          // fill telegramm header - just for later debugging ( the header is part of the command payload itselfy ) {{{
          Telegram.PlcToRob.Sequence[_seqIdx].Fragment[_fragIdx].Command.Header.CmdType       := CombineBytesToUint ( AxesGroup.Acyclic.ActiveCommandRegister.Register[_regIdx].Command[ACTIVE_CMD].Payload[0],
                                                                                                                      AxesGroup.Acyclic.ActiveCommandRegister.Register[_regIdx].Command[ACTIVE_CMD].Payload[1]);
          Telegram.PlcToRob.Sequence[_seqIdx].Fragment[_fragIdx].Command.Header.ExecMode.0    :=                      AxesGroup.Acyclic.ActiveCommandRegister.Register[_regIdx].Command[ACTIVE_CMD].Payload[2].0;
          Telegram.PlcToRob.Sequence[_seqIdx].Fragment[_fragIdx].Command.Header.ExecMode.1    :=                      AxesGroup.Acyclic.ActiveCommandRegister.Register[_regIdx].Command[ACTIVE_CMD].Payload[2].1;
          Telegram.PlcToRob.Sequence[_seqIdx].Fragment[_fragIdx].Command.Header.ExecMode.2    :=                      AxesGroup.Acyclic.ActiveCommandRegister.Register[_regIdx].Command[ACTIVE_CMD].Payload[2].2;
          Telegram.PlcToRob.Sequence[_seqIdx].Fragment[_fragIdx].Command.Header.ExecMode.3    :=                      AxesGroup.Acyclic.ActiveCommandRegister.Register[_regIdx].Command[ACTIVE_CMD].Payload[2].3;
          Telegram.PlcToRob.Sequence[_seqIdx].Fragment[_fragIdx].Command.Header.Prio.0        :=                      AxesGroup.Acyclic.ActiveCommandRegister.Register[_regIdx].Command[ACTIVE_CMD].Payload[3].0;
          Telegram.PlcToRob.Sequence[_seqIdx].Fragment[_fragIdx].Command.Header.Prio.1        :=                      AxesGroup.Acyclic.ActiveCommandRegister.Register[_regIdx].Command[ACTIVE_CMD].Payload[3].1;
          Telegram.PlcToRob.Sequence[_seqIdx].Fragment[_fragIdx].Command.Header.Prio.2        :=                      AxesGroup.Acyclic.ActiveCommandRegister.Register[_regIdx].Command[ACTIVE_CMD].Payload[3].2;
          Telegram.PlcToRob.Sequence[_seqIdx].Fragment[_fragIdx].Command.Header.Prio.3        :=                      AxesGroup.Acyclic.ActiveCommandRegister.Register[_regIdx].Command[ACTIVE_CMD].Payload[3].3;
          Telegram.PlcToRob.Sequence[_seqIdx].Fragment[_fragIdx].Command.Header.ParSequence.0 :=                      AxesGroup.Acyclic.ActiveCommandRegister.Register[_regIdx].Command[ACTIVE_CMD].Payload[3].4;
          Telegram.PlcToRob.Sequence[_seqIdx].Fragment[_fragIdx].Command.Header.ParSequence.1 :=                      AxesGroup.Acyclic.ActiveCommandRegister.Register[_regIdx].Command[ACTIVE_CMD].Payload[3].5;
          Telegram.PlcToRob.Sequence[_seqIdx].Fragment[_fragIdx].Command.Header.ParSequence.2 :=                      AxesGroup.Acyclic.ActiveCommandRegister.Register[_regIdx].Command[ACTIVE_CMD].Payload[3].6;
          Telegram.PlcToRob.Sequence[_seqIdx].Fragment[_fragIdx].Command.Header.ParSequence.3 :=                      AxesGroup.Acyclic.ActiveCommandRegister.Register[_regIdx].Command[ACTIVE_CMD].Payload[3].7;
          // }}}
          // loop through the payload
          FOR _payLoadPtr := AxesGroup.Acyclic.ActiveCommandRegister.Register[_regIdx].Command[ACTIVE_CMD].PayLoadPtr TO AxesGroup.Acyclic.ActiveCommandRegister.Register[_regIdx].Command[ACTIVE_CMD].PayloadLen -1  
          DO
            // copy payload
            Telegram.PlcToRob.Sequence[_seqIdx].Fragment[_fragIdx].Command.Payload[_payLoadPtr] 
              := AxesGroup.Acyclic.ActiveCommandRegister.Register[_regIdx].Command[ACTIVE_CMD].Payload[_payLoadPtr];
        
            // inc current sequence payload length
            Telegram.PlcToRob.Sequence[_seqIdx].Header.PayloadLength
              := Telegram.PlcToRob.Sequence[_seqIdx].Header.PayloadLength + 1;  
        
            // inc current fragment payload length
            Telegram.PlcToRob.Sequence[_seqIdx].Fragment[_fragIdx].Header.PayloadLength 
              := Telegram.PlcToRob.Sequence[_seqIdx].Fragment[_fragIdx].Header.PayloadLength + 1;
        
            // inc payload pointer in active command register
            AxesGroup.Acyclic.ActiveCommandRegister.Register[_regIdx].Command[ACTIVE_CMD].PayLoadPtr 
              := AxesGroup.Acyclic.ActiveCommandRegister.Register[_regIdx].Command[ACTIVE_CMD].PayLoadPtr + 1;
          
            // set command state
            IF ( AxesGroup.Acyclic.ActiveCommandRegister.Register[_regIdx].Command[ACTIVE_CMD].PayLoadPtr >= AxesGroup.Acyclic.ActiveCommandRegister.Register[_regIdx].Command[ACTIVE_CMD].PayLoadLen) 
            THEN
              AxesGroup.Acyclic.ActiveCommandRegister.Register[_regIdx].Command[ACTIVE_CMD].State := BufferStateCmd.PROCESSED;
            ELSE
              AxesGroup.Acyclic.ActiveCommandRegister.Register[_regIdx].Command[ACTIVE_CMD].State := BufferStateCmd.SENDING;  
            END_IF 
    
            // calc current telegram payload length
           _telegramLengthCurrent := 4 + Telegram.PlcToRob.Sequence[_seqIdx].Header.PayloadLength; // ST-FIX F63: sequence header + payload
      
            // check limit reached ?
            IF ( _telegramLengthCurrent >= SEQUENCE_MAX_PAYLOAD_SIZE (* ST-FIX F63 *)) 
            THEN  
              EXIT; // -> abort for loop 
            END_IF  
          END_FOR
    
          // check payload complete ?
         _fragmentAction.Complete := AxesGroup.Acyclic.ActiveCommandRegister.Register[_regIdx].Command[ACTIVE_CMD].PayLoadPtr 
                                  >= AxesGroup.Acyclic.ActiveCommandRegister.Register[_regIdx].Command[ACTIVE_CMD].PayloadLen;
    
          // just for brakepoint
          IF (_fragmentAction.Complete)
          THEN
           _fragmentAction.Complete := _fragmentAction.Complete; 
          END_IF
    
          // set fragment action
          Telegram.PlcToRob.Sequence[_seqIdx].Fragment[_fragIdx].Header.FragmentAction := FragmentActionToByte(_fragmentAction);
        END_IF
      END_IF
      
      // inc execution order list index 
     _listIdx := _listIdx + 1;
      // inc fragment index 
     _fragIdx := _fragIdx + 1;
  
      // check abort conditions
      IF (( _telegramLengthCurrent                                                >= SEQUENCE_MAX_PAYLOAD_SIZE (* ST-FIX F63 *)  ) OR  // Payload limit reached 
          ( _fragIdx                                                              >=  RobotLibraryParameter.FRAGMENT_MAX ) OR  // Max fragment limit reached
          (  AxesGroup.Acyclic.ActiveCommandRegister.ExecutionOrderList[_listIdx]  =  EMPTY_EOL_ENTRY                    ))    // No entry in ExecutionOrderList left
      THEN
        EXIT;// -> Abort while loop
      END_IF         
    END_WHILE  
    
    AxesGroup.State.SequenceCountSend          := _seqCount; // ST-FIX F63
    AxesGroup.State.FragmentCountSend[_seqIdx] := _fragIdx;
    
  END_IF  
END_FOR
                
                
END_METHOD

METHOD CalculateCyclicDataLength : UINT
VAR_IN_OUT
  /// Robot assignment of function
  AxesGroup : AxesGroup;
END_VAR
VAR_INPUT
  /// Communication direction
  Direction : ComDirection;
END_VAR

VAR CONSTANT
  /// Size of the header
  ROB_TO_PLC_HEADER_SIZE : UINT := 10;
END_VAR
                  // ------------------------------------
// PLC -> ROB
// ------------------------------------
IF (Direction = ComDirection.PLC_TO_ROB)
THEN  
  // Add Header size 
  CalculateCyclicDataLength := CalculateCyclicDataLength + SIZEOF(Telegram.PlcToRob.Header);  
  // Add Cyclic size (ST-FIX F2: only with Cartesian Position RC -> PLC)
  IF ( AxesGroup.CyclicOptional.RobToPlc.CartesianPosition.Active )
  THEN
    CalculateCyclicDataLength := CalculateCyclicDataLength + SIZEOF(Telegram.PlcToRob.Cyclic);
  END_IF
  
  // Check SubProgramData active ? 
  IF ( AxesGroup.CyclicOptional.PlcToRob.SubProgramData.Active )
  THEN
    // Add SubProgramData size 
    CalculateCyclicDataLength := CalculateCyclicDataLength + SIZEOF(Telegram.PlcToRob.CyclicOptional.SubProgramData);
  END_IF
    
  // Check CartesianPosition active ? 
  IF ( AxesGroup.CyclicOptional.PlcToRob.CartesianPosition.Active )
  THEN
    // Add CartesianPosition size 
    CalculateCyclicDataLength := CalculateCyclicDataLength + SIZEOF(Telegram.PlcToRob.CyclicOptional.CartesianPosition);
  END_IF
  
  // Check JointPosition active ? 
  IF ( AxesGroup.CyclicOptional.PlcToRob.JointPosition.Active )
  THEN
    // Add JointPosition size 
    CalculateCyclicDataLength := CalculateCyclicDataLength + SIZEOF(Telegram.PlcToRob.CyclicOptional.JointPosition);
  END_IF  
  
  // Check Force active ? 
  IF ( AxesGroup.CyclicOptional.PlcToRob.Force.Active )
  THEN
    // Add Force size 
    CalculateCyclicDataLength := CalculateCyclicDataLength + SIZEOF(Telegram.PlcToRob.CyclicOptional.Force);
  END_IF  
    
  // Check CartesianPositionExt acive ? 
  IF ( AxesGroup.CyclicOptional.PlcToRob.CartesianPositionExt.Active )
  THEN
    // Add CartesianPositionExt size 
    CalculateCyclicDataLength := CalculateCyclicDataLength + SIZEOF(Telegram.PlcToRob.CyclicOptional.CartesianPositionExt);
  END_IF   
    
  // Check JointPositionExt active ?
  IF ( AxesGroup.CyclicOptional.PlcToRob.JointPositionExt.Active )
  THEN
    // Add JointPositionExt size 
    CalculateCyclicDataLength := CalculateCyclicDataLength + SIZEOF(Telegram.PlcToRob.CyclicOptional.JointPositionExt);
  END_IF  
        
  // Check ForceExt active ?
  IF ( AxesGroup.CyclicOptional.PlcToRob.ForceExt.Active )
  THEN
    // Add ForceExt size 
    CalculateCyclicDataLength := CalculateCyclicDataLength + SIZEOF(Telegram.PlcToRob.CyclicOptional.ForceExt);
  END_IF
END_IF

// ------------------------------------
// ROB -> PLC
// ------------------------------------
IF (Direction = ComDirection.ROB_TO_PLC)
THEN
  // Add Header size 
  CalculateCyclicDataLength := CalculateCyclicDataLength + ROB_TO_PLC_HEADER_SIZE; 
  // a constant, because SIZEOF(Telegram.RobToPlc.Header) counts the VersionStruct instead of one byte
  
  // Check SubProgramData active ? 
  IF ( AxesGroup.CyclicOptional.RobToPlc.SubProgramData.Active )
  THEN
    // Add SubProgramData size 
    CalculateCyclicDataLength := CalculateCyclicDataLength + SIZEOF(Telegram.RobToPlc.CyclicOptional.SubProgramData);
  END_IF
    
  // Check CartesianPosition active ? 
  IF ( AxesGroup.CyclicOptional.RobToPlc.CartesianPosition.Active )
  THEN
    // Add CartesianPosition size 
    CalculateCyclicDataLength := CalculateCyclicDataLength + SIZEOF(Telegram.RobToPlc.CyclicOptional.CartesianPosition);
  END_IF
  
  // Check JointPosition active ? 
  IF ( AxesGroup.CyclicOptional.RobToPlc.JointPosition.Active )
  THEN
    // Add JointPosition size 
    CalculateCyclicDataLength := CalculateCyclicDataLength + SIZEOF(Telegram.RobToPlc.CyclicOptional.JointPosition);
  END_IF  
  
  // Check Force active ? 
  IF ( AxesGroup.CyclicOptional.RobToPlc.Force.Active )
  THEN
    // Add Force size 
    CalculateCyclicDataLength := CalculateCyclicDataLength + SIZEOF(Telegram.RobToPlc.CyclicOptional.Force);
  END_IF  
    
  // Check Current acive ? 
  IF ( AxesGroup.CyclicOptional.RobToPlc.Current.Active )
  THEN
    // Add Current size 
    CalculateCyclicDataLength := CalculateCyclicDataLength + SIZEOF(Telegram.RobToPlc.CyclicOptional.Current);
  END_IF    
    
  // Check CartesianPositionExt acive ? 
  IF ( AxesGroup.CyclicOptional.RobToPlc.CartesianPositionExt.Active )
  THEN
    // Add CartesianPositionExt size 
    CalculateCyclicDataLength := CalculateCyclicDataLength + SIZEOF(Telegram.RobToPlc.CyclicOptional.CartesianPositionExt);
  END_IF  
    
  // Check JointPositionExt active ?
  IF ( AxesGroup.CyclicOptional.RobToPlc.JointPositionExt.Active )
  THEN
    // Add JointPositionExt size 
    CalculateCyclicDataLength := CalculateCyclicDataLength + SIZEOF(Telegram.RobToPlc.CyclicOptional.JointPositionExt);
  END_IF  
        
  // Check ForceExt active ?
  IF ( AxesGroup.CyclicOptional.RobToPlc.ForceExt.Active )
  THEN
    // Add ForceExt size 
    CalculateCyclicDataLength := CalculateCyclicDataLength + SIZEOF(Telegram.RobToPlc.CyclicOptional.ForceExt);
  END_IF
    
  // Check CurrentExt active ? 
  IF ( AxesGroup.CyclicOptional.RobToPlc.CurrentExt.Active )
  THEN
    // Add CurrentExt size 
    CalculateCyclicDataLength := CalculateCyclicDataLength + SIZEOF(Telegram.RobToPlc.CyclicOptional.CurrentExt);
  END_IF
END_IF
                
END_METHOD

METHOD CalculateSequencePayloadMax : UINT
VAR_IN_OUT
  /// Robot assignment of function
  AxesGroup : AxesGroup;
END_VAR
VAR_INPUT
  /// Communication direction
  Direction : ComDirection;
  /// Sequeunce
  Sequence : SequenceFlag;  
END_VAR

VAR
  /// Length of the cyclic header
 _cyclicDataLength      : UINT;
  /// Acyclic area (ST-FIX F63)
 _area                  : UDINT;
END_VAR
                  // calculate cyclic header length
_cyclicDataLength := CalculateCyclicDataLength(AxesGroup := AxesGroup, Direction := Direction);


// ST-FIX F63: acyclic area without the footer, halved for two sequences (spec Fig. 5-205)
IF ( Direction = ComDirection.PLC_TO_ROB )
THEN
  _area := UINT_TO_UDINT(_parCfg.Com.TelegramLengthPlcToRob) - UINT_TO_UDINT(_cyclicDataLength) - FOOTER_SIZE;
ELSE
  _area := UINT_TO_UDINT(_parCfg.Com.TelegramLengthRobToPlc) - UINT_TO_UDINT(_cyclicDataLength) - FOOTER_SIZE;
END_IF

IF ( NOT _parCfg.Com.TwoSequences )
THEN
  IF ( Sequence = SequenceFlag.PRIMARY_SEQUENCE )
  THEN
    CalculateSequencePayloadMax := UDINT_TO_UINT(_area);
  ELSE
    CalculateSequencePayloadMax := 0;
  END_IF
ELSIF ( Sequence = SequenceFlag.PRIMARY_SEQUENCE )
THEN
  CalculateSequencePayloadMax := UDINT_TO_UINT(_area / 2);
ELSE
  CalculateSequencePayloadMax := UDINT_TO_UINT(_area - _area / 2);
END_IF
                
END_METHOD

METHOD CalculateSequencePayloadStartAdr : UINT
VAR_IN_OUT
  /// Robot assignment of function
  AxesGroup : AxesGroup;
END_VAR
VAR_INPUT
  /// Communication direction
  Direction : ComDirection;
  /// Sequeunce
  Sequence : SequenceFlag;  
END_VAR

VAR
  /// Length of the cyclic header
 _cyclicDataLength      : UINT;
  /// Length of the sequnce payload
 _sequencePayloadLength : UINT;
END_VAR
                  // calculate cyclic header length
_cyclicDataLength := CalculateCyclicDataLength(AxesGroup := AxesGroup, Direction := Direction);

CASE (Sequence) 
OF

  SequenceFlag.PRIMARY_SEQUENCE   : 
  
    // return start address
    CalculateSequencePayloadStartAdr := _cyclicDataLength;

  SequenceFlag.SECONDARY_SEQUENCE :
  
    // calculate sequence payload max
   _sequencePayloadLength 
     := CalculateSequencePayloadMax( AxesGroup := AxesGroup, 
                                     Direction := Direction, 
                                     Sequence  := SequenceFlag.PRIMARY_SEQUENCE ); // ST-FIX F63: behind the area of the 1st sequence
                                     
    // return start address
    CalculateSequencePayloadStartAdr := _cyclicDataLength + _sequencePayloadLength;
    
END_CASE
                
END_METHOD

METHOD PROTECTED CalculateTelegramLengthPlcToRob : UINT
VAR_IN_OUT
  /// Robot assignment of function
  AxesGroup : AxesGroup;
END_VAR
VAR
  /// length of the cyclic data block
 _cyclicDataLength : UINT;
END_VAR
                  _cyclicDataLength := CalculateCyclicDataLength(AxesGroup := AxesGroup, Direction := ComDirection.PLC_TO_ROB); 


IF ( _parCfg.Com.TwoSequences )
THEN
  CalculateTelegramLengthPlcToRob := _cyclicDataLength
                                    + SIZEOF(Telegram.PlcToRob.Sequence[  PRIMARY_SEQUENCE].Header)
                                    +       (Telegram.PlcToRob.Sequence[  PRIMARY_SEQUENCE].Header.PayloadLength)
                                    + SIZEOF(Telegram.PlcToRob.Sequence[SECONDARY_SEQUENCE].Header)
                                    +       (Telegram.PlcToRob.Sequence[SECONDARY_SEQUENCE].Header.PayloadLength)
                                    + SIZEOF(Telegram.PlcToRob.Footer);  
ELSE
  CalculateTelegramLengthPlcToRob := _cyclicDataLength
                                    + SIZEOF(Telegram.PlcToRob.Sequence[PRIMARY_SEQUENCE].Header)
                                    +       (Telegram.PlcToRob.Sequence[PRIMARY_SEQUENCE].Header.PayloadLength)
                                    + SIZEOF(Telegram.PlcToRob.Footer);
END_IF
                
END_METHOD

/// ST-FIX F132: checks that the AxesGroup and the telegram buffers are not used by another RobotTask
/// (table 7-1: 16#8007 ERR_AXESGROUP_INVALID, 16#8008 ERR_PERIPHERY_INVALID) and registers them
METHOD PRIVATE CheckAssignmentValid : BOOL
VAR_IN_OUT
  /// Robot assignment of function
  AxesGroup    : AxesGroup;
  /// Inputs of PLC for communication from RC
  RobotInData  : ARRAY[*] OF BYTE;
  /// Outputs of PLC for communication to RC
  RobotOutData : ARRAY[*] OF BYTE;
END_VAR
VAR
  /// Loop index over the entries
 _idx     : DINT;
  /// Entry of this instance
 _own     : DINT;
  /// First free entry
 _free    : DINT;
  /// Address of RobotInData
 _inAdr   : PVOID;
  /// Address of RobotOutData
 _outAdr  : PVOID;
END_VAR
                  CheckAssignmentValid := FALSE;

// AxesGroup used by another RobotTask ?
IF (( AxesGroup.State.RobotTaskId <> 0           ) AND
    ( AxesGroup.State.RobotTaskId <> _instanceId ))
THEN
  IF ( ErrorID <> RobotLibraryErrorIdEnum.ERR_AXESGROUP_INVALID )
  THEN
    SetError( ErrorID := RobotLibraryErrorIdEnum.ERR_AXESGROUP_INVALID, Overwrite := TRUE );
    // Create log entry
    CreateLogMessagePara1 ( Timestamp   := SystemTime,
                            MessageType := MessageType.CMD,
                            Severity    := Severity.ERROR,
                            MessageCode := ErrorID,
                            MessageText := 'AxesGroup is already used by RobotTask {1}',
                            Para1       := UDINT_TO_STRING(AxesGroup.State.RobotTaskId));
  END_IF
  RETURN;
END_IF

// telegram buffers used by another RobotTask ?
_inAdr  := ADR(RobotInData [ROBOT_IN_DATA_MIN ]);
_outAdr := ADR(RobotOutData[ROBOT_OUT_DATA_MIN]);
_own    := 0;
_free   := 0;
FOR _idx := 1 TO PERIPHERY_ENTRIES
DO
  IF ( _peripheryOwner[_idx] = _instanceId )
  THEN
   _own := _idx;
  ELSIF ( _peripheryOwner[_idx] = 0 )
  THEN
    IF ( _free = 0 )
    THEN
     _free := _idx;
    END_IF
  ELSIF (( _peripheryInAdr [_idx] = _inAdr  ) OR
         ( _peripheryOutAdr[_idx] = _outAdr ))
  THEN
    IF ( ErrorID <> RobotLibraryErrorIdEnum.ERR_PERIPHERY_INVALID )
    THEN
      SetError( ErrorID := RobotLibraryErrorIdEnum.ERR_PERIPHERY_INVALID, Overwrite := TRUE );
      // Create log entry
      CreateLogMessagePara1 ( Timestamp   := SystemTime,
                              MessageType := MessageType.CMD,
                              Severity    := Severity.ERROR,
                              MessageCode := ErrorID,
                              MessageText := 'Telegram buffers are already used by RobotTask {1}',
                              Para1       := UDINT_TO_STRING(_peripheryOwner[_idx]));
    END_IF
    RETURN;
  END_IF
END_FOR

// register this instance (the addresses can change after an online change)
IF ( _own = 0 )
THEN
 _own := _free;
END_IF
IF ( _own > 0 )
THEN
 _peripheryOwner [_own] := _instanceId;
 _peripheryInAdr [_own] := _inAdr;
 _peripheryOutAdr[_own] := _outAdr;
END_IF
AxesGroup.State.RobotTaskId := _instanceId;

CheckAssignmentValid := TRUE;
                
END_METHOD

METHOD PROTECTED CheckParameterChanged : BOOL
VAR_IN_OUT
  /// Robot assignment of function
  AxesGroup    : AxesGroup; 
END_VAR

VAR
  /// internal index for loops
 _idx : DINT;
END_VAR
                  // Check initialization is already done ?
IF ( NOT Initialized )
THEN
  CheckParameterChanged := FALSE;
  RETURN;
END_IF

// compare memory 
CheckParameterChanged := ( SysDepMemCmp(pData1 := ADR(ParCfg), pData2 := ADR(_parCfg), DataLen := SIZEOF(ParCfg)) <> RobotLibraryConstants.OK );

FOR _idx := SyncTime.DURING_START_UP TO SyncTime.AFTER_START_UP
DO
  // Check Tool SyncMode changed ? 
  IF ( _parCfg.Plc.Parameter.SynchronizationModes.Tool[_idx] <> ParCfg.Plc.Parameter.SynchronizationModes.Tool[_idx] )
  THEN
    // Set info
    SetInfo( InfoID := RobotLibraryInfoIdEnum.INFO_CHANGE_TOOL_SYNC_MODE_TO_NEGATIVE_ONLY_AT_PLC_START_ALLOWED, Overwrite := TRUE);
     
    // Create log entry
    CreateLogMessagePara3( Timestamp   := SystemTime,
                           MessageType := MessageType.CMD,
                           Severity    := Severity.INFO,
                           MessageCode := 0,
                           MessageText := 'SyncMode.Tool[{1}] changed from {2} to {3}, but this is only allowed at PLC start',
                           Para1       := SYNC_TIME_TO_STRING(_idx),
                           Para2       := SYNC_MODE_TO_STRING( ParCfg.Plc.Parameter.SynchronizationModes.Tool[_idx]),
                           Para3       := SYNC_MODE_TO_STRING(_parCfg.Plc.Parameter.SynchronizationModes.Tool[_idx]));   
  END_IF
  
  
  // Check Frame SyncMode changed ? 
  IF ( _parCfg.Plc.Parameter.SynchronizationModes.Frame[_idx] <> ParCfg.Plc.Parameter.SynchronizationModes.Frame[_idx] )
  THEN
    // Set info
    SetInfo( InfoID := RobotLibraryInfoIdEnum.INFO_CHANGE_FRAME_SYNC_MODE_TO_NEGATIVE_ONLY_AT_PLC_START_ALLOWED, Overwrite :=  TRUE);
     
    // Create log entry
    CreateLogMessagePara3( Timestamp   := SystemTime,
                           MessageType := MessageType.CMD,
                           Severity    := Severity.INFO,
                           MessageCode := 0,
                           MessageText := 'SyncMode.Frame[{1}] changed from {2} to {3}, but this is only allowed at PLC start',
                           Para1       := SYNC_TIME_TO_STRING(_idx),
                           Para2       := SYNC_MODE_TO_STRING( ParCfg.Plc.Parameter.SynchronizationModes.Frame[_idx]),
                           Para3       := SYNC_MODE_TO_STRING(_parCfg.Plc.Parameter.SynchronizationModes.Frame[_idx]));   
  END_IF
  
  
  // Check Load SyncMode changed ? 
  IF ( _parCfg.Plc.Parameter.SynchronizationModes.Load[_idx] <> ParCfg.Plc.Parameter.SynchronizationModes.Load[_idx] )
  THEN
    // Set info
    SetInfo( InfoID := RobotLibraryInfoIdEnum.INFO_CHANGE_LOAD_SYNC_MODE_TO_NEGATIVE_ONLY_AT_PLC_START_ALLOWED, Overwrite := TRUE);
     
    // Create log entry
    CreateLogMessagePara3( Timestamp   := SystemTime,
                           MessageType := MessageType.CMD,
                           Severity    := Severity.INFO,
                           MessageCode := 0,
                           MessageText := 'SyncMode.Load[{1}] changed from {2} to {3}, but this is only allowed at PLC start',
                           Para1       := SYNC_TIME_TO_STRING(_idx),
                           Para2       := SYNC_MODE_TO_STRING( ParCfg.Plc.Parameter.SynchronizationModes.Load[_idx]),
                           Para3       := SYNC_MODE_TO_STRING(_parCfg.Plc.Parameter.SynchronizationModes.Load[_idx]));   
  END_IF
  
  
  // Check WorkAreas SyncMode changed ? 
  IF ( _parCfg.Plc.Parameter.SynchronizationModes.WorkAreas[_idx] <> ParCfg.Plc.Parameter.SynchronizationModes.WorkAreas[_idx] )
  THEN
    // Set info
    SetInfo( InfoID := RobotLibraryInfoIdEnum.INFO_CHANGE_WORK_AREA_SYNC_MODE_TO_NEGATIVE_ONLY_AT_PLC_START_ALLOWED, Overwrite := TRUE);
     
    // Create log entry
    CreateLogMessagePara3( Timestamp   := SystemTime,
                           MessageType := MessageType.CMD,
                           Severity    := Severity.INFO,
                           MessageCode := 0,
                           MessageText := 'SyncMode.WorkAreas[{1}] changed from {2} to {3}, but this is only allowed at PLC start',
                           Para1       := SYNC_TIME_TO_STRING(_idx),
                           Para2       := SYNC_MODE_TO_STRING( ParCfg.Plc.Parameter.SynchronizationModes.WorkAreas[_idx]),
                           Para3       := SYNC_MODE_TO_STRING(_parCfg.Plc.Parameter.SynchronizationModes.WorkAreas[_idx]));   
  END_IF

  // Check SWLimits SyncMode changed ? 
  IF ( _parCfg.Plc.Parameter.SynchronizationModes.SWLimits[_idx] <> ParCfg.Plc.Parameter.SynchronizationModes.SWLimits[_idx] )
  THEN
    // Set info
    SetInfo( InfoID := RobotLibraryInfoIdEnum.INFO_CHANGE_SWLIMITS_SYNC_MODE_TO_NEGATIVE_ONLY_AT_PLC_START_ALLOWED, Overwrite := TRUE);
     
    // Create log entry
    CreateLogMessagePara3( Timestamp   := SystemTime,
                           MessageType := MessageType.CMD,
                           Severity    := Severity.INFO,
                           MessageCode := 0,
                           MessageText := 'SyncMode.SWLimits[{1}] changed from {2} to {3}, but this is only allowed at PLC start',
                           Para1       := SYNC_TIME_TO_STRING(_idx),
                           Para2       := SYNC_MODE_TO_STRING( ParCfg.Plc.Parameter.SynchronizationModes.SWLimits[_idx]),
                           Para3       := SYNC_MODE_TO_STRING(_parCfg.Plc.Parameter.SynchronizationModes.SWLimits[_idx]));   
  END_IF
  
 
  // Check DefaultDynamics SyncMode changed ? 
  IF ( _parCfg.Plc.Parameter.SynchronizationModes.DefaultDynamics[_idx] <> ParCfg.Plc.Parameter.SynchronizationModes.DefaultDynamics[_idx] )
  THEN
    // Set info
    SetInfo( InfoID := RobotLibraryInfoIdEnum.INFO_CHANGE_DEFAULT_DYNAMICS_SYNC_MODE_TO_NEGATIVE_ONLY_AT_PLC_START_ALLOWED, Overwrite := TRUE);
     
    // Create log entry
    CreateLogMessagePara3( Timestamp   := SystemTime,
                           MessageType := MessageType.CMD,
                           Severity    := Severity.INFO,
                           MessageCode := 0,
                           MessageText := 'SyncMode.DefaultDynamics[{1}] changed from {2} to {3}, but this is only allowed at PLC start',
                           Para1       := SYNC_TIME_TO_STRING(_idx),
                           Para2       := SYNC_MODE_TO_STRING( ParCfg.Plc.Parameter.SynchronizationModes.DefaultDynamics[_idx]),
                           Para3       := SYNC_MODE_TO_STRING(_parCfg.Plc.Parameter.SynchronizationModes.DefaultDynamics[_idx]));   
  END_IF
  
  
  // Check ReferenceDynamics SyncMode changed ?
  IF ( _parCfg.Plc.Parameter.SynchronizationModes.ReferenceDynamics[_idx] <> ParCfg.Plc.Parameter.SynchronizationModes.ReferenceDynamics[_idx] )
  THEN
    // Set info
    SetInfo(InfoID := RobotLibraryInfoIdEnum.INFO_CHANGE_REFERENCE_DYNAMICS_SYNC_MODE_TO_NEGATIVE_ONLY_AT_PLC_START_ALLOWED, Overwrite := TRUE );
     
    // Create log entry
    CreateLogMessagePara3( Timestamp   := SystemTime,
                           MessageType := MessageType.CMD,
                           Severity    := Severity.INFO,
                           MessageCode := 0,
                           MessageText := 'SyncMode.ReferenceDynamics[{1}] changed from {2} to {3}, but this is only allowed at PLC start',
                           Para1       := SYNC_TIME_TO_STRING(_idx),
                           Para2       := SYNC_MODE_TO_STRING( ParCfg.Plc.Parameter.SynchronizationModes.ReferenceDynamics[_idx]),
                           Para3       := SYNC_MODE_TO_STRING(_parCfg.Plc.Parameter.SynchronizationModes.ReferenceDynamics[_idx]));   
  END_IF

END_FOR


// Check Plc.OptionalCyclic changed ? 
IF ( PlcOptionalCyclicToUint(_parCfg.Plc.OptionalCyclic) <> PlcOptionalCyclicToUint(ParCfg.Plc.OptionalCyclic ))
THEN
  // Set error
  SetWarning( WarningID := RobotLibraryWarningIdEnum.WARN_TELEGRAM_NO_CHANGED_DURING_OPERATION, Overwrite := TRUE ); // ST-FIX F68
   
  // Create log entry
  CreateLogMessagePara2( Timestamp   := SystemTime,
                         MessageType := MessageType.CMD,
                         Severity    := Severity.WARNING,
                         MessageCode := 0,
                         MessageText := 'ParCfg.Plc.OptionalCyclic changed after initialization from {1} to {2} -> Reinitialize by disabling and enabling the RobotTask',
                         Para1       := WORD_TO_STRING_BIN(PlcOptionalCyclicToUint(_parCfg.Plc.OptionalCyclic)),
                         Para2       := WORD_TO_STRING_BIN(PlcOptionalCyclicToUint( ParCfg.Plc.OptionalCyclic)));   
END_IF


// Check Rob.OptionalCyclic changed ? 
IF ( RobOptionalCyclicToUint(_parCfg.Rob.OptionalCyclic) <> RobOptionalCyclicToUint(ParCfg.Rob.OptionalCyclic ))
THEN
  // Set error
  SetWarning( WarningID := RobotLibraryWarningIdEnum.WARN_TELEGRAM_NO_CHANGED_DURING_OPERATION, Overwrite := TRUE ); // ST-FIX F68
   
  // Create log entry
  CreateLogMessagePara2( Timestamp   := SystemTime,
                         MessageType := MessageType.CMD,
                         Severity    := Severity.WARNING,
                         MessageCode := 0,
                         MessageText := 'ParCfg.Rob.OptionalCyclic changed after initialization from {1} to {2} -> Reinitialize by disabling and enabling the RobotTask',
                         Para1       := WORD_TO_STRING_BIN(RobOptionalCyclicToUint(_parCfg.Rob.OptionalCyclic)),
                         Para2       := WORD_TO_STRING_BIN(RobOptionalCyclicToUint( ParCfg.Rob.OptionalCyclic)));   
END_IF

                
                
END_METHOD

METHOD PROTECTED CheckParameterValid : BOOL
VAR_IN_OUT
  /// Robot assignment of function
  AxesGroup : AxesGroup; 
END_VAR
                  // init return value
CheckParameterValid := TRUE;


// Check ParCfg.Com.TelegramLengthPlcToRob
IF ( ParCfg.Com.TelegramLengthPlcToRob < 128 )
THEN
  // Set Warning
  SetWarning( WarningID := RobotLibraryWarningIdEnum.WARN_ACYCLIC_RANGE_PLC_TO_ROB_VERY_SMALL, Overwrite := TRUE );
END_IF

// Check ParCfg.Com.TelegramLengthRobToPlc
IF ( ParCfg.Com.TelegramLengthRobToPlc < 128 )
THEN
  // Set Warning
  SetWarning( WarningID := RobotLibraryWarningIdEnum.WARN_ACYCLIC_RANGE_ROB_TO_PLC_VERY_SMALL, Overwrite := TRUE );
END_IF



// Region ParCfg.Com {{{

// Check LifeSignTimeout
IF ( ParCfg.Com.LifeSignTimeOut < T#10MS )
THEN
  // set to valid min value
  ParCfg.Com.LifeSignTimeOut := T#10MS;
 
  // Set info
  SetInfo( InfoID := RobotLibraryInfoIdEnum.INFO_LIFESIGN_TIMEOUT_TO_SMALL_AND_SET_TO_10MS, Overwrite := TRUE);
   
  // Create log entry
  CreateLogMessagePara1 ( Timestamp   := SystemTime,
                          MessageType := MessageType.CMD,
                          Severity    := Severity.INFO,
                          MessageCode := 0,
                          MessageText := 'LifeSignTimeout to small and set from {1}ms to 10ms',
                          Para1       := TIME_TO_STRING(ParCfg.Com.LifeSignTimeOut));                          
END_IF


// Check ParCfg.Com.TelegramLengthPlcToRob
IF (( ParCfg.Com.TelegramLengthPlcToRob < 64                  ) OR
    ( ParCfg.Com.TelegramLengthPlcToRob > ROBOT_OUT_DATA_SIZE ))
THEN
  // parameter(s) not valid
  CheckParameterValid := FALSE;

  // Set error
  SetError( ErrorID := RobotLibraryErrorIdEnum.ERR_TELEGRAM_LENGTH_MISMATCH_0x80A3, Overwrite := TRUE );
   
  // Create log entry
  CreateLogMessagePara1 ( Timestamp   := SystemTime,
                          MessageType := MessageType.CMD,
                          Severity    := Severity.INFO,
                          MessageCode := 0,
                          MessageText :=               'ParCfg.Com.TelegramLengthPlcToRob {1} invalid',
                          Para1       := UINT_TO_STRING(ParCfg.Com.TelegramLengthPlcToRob));
  // no further validation                          
  RETURN;                          
END_IF

// Check ParCfg.Com.TelegramLengthRobToPlc
IF (( ParCfg.Com.TelegramLengthRobToPlc < 64                 ) OR
    ( ParCfg.Com.TelegramLengthRobToPlc > ROBOT_IN_DATA_SIZE ))
THEN
  // parameter(s) not valid
  CheckParameterValid := FALSE;

  // Set error
  SetError( ErrorID := RobotLibraryErrorIdEnum.ERR_TELEGRAM_LENGTH_MISMATCH_0x80A3, Overwrite := TRUE );
   
  // Create log entry
  CreateLogMessagePara1 ( Timestamp   := SystemTime,
                          MessageType := MessageType.CMD,
                          Severity    := Severity.INFO,
                          MessageCode := 0,
                          MessageText :=               'ParCfg.Com.TelegramLengthRobToPlc {1} invalid',
                          Para1       := UINT_TO_STRING(ParCfg.Com.TelegramLengthRobToPlc));
  // no further validation                          
  RETURN;                          
END_IF
// ST-FIX F63: two telegram sequences must be activated in both directions and for the layout
IF ( ParCfg.Plc.OptionalCyclic.UseTwoSequences <> ParCfg.Rob.OptionalCyclic.UseTwoSequences ) OR
   ( ParCfg.Plc.OptionalCyclic.UseTwoSequences <> ParCfg.Com.TwoSequences                  )
THEN
  CheckParameterValid := FALSE;
  SetError( ErrorID := RobotLibraryErrorIdEnum.ERR_TELEGRAM_NUMBER_INVALID_0x80AB, Overwrite := TRUE );
  CreateLogMessage( Timestamp   := SystemTime,
                    MessageType := MessageType.CMD,
                    Severity    := Severity.ERROR,
                    MessageCode := 0,
                    MessageText := 'TwoSequences must be set in Com and in Plc/Rob.OptionalCyclic');
  RETURN;
END_IF
// EndRegion }}}

// Region ParCfg.Rob.OptionalCyclic {{{

// Check configuration if optional cyclic CartesianPosition valid ?
// ST-FIX F137: the extended cartesian position cannot be used without the cartesian position ->
// the cartesian position is activated automatically (spec 6.4.2 and InfoID 16#6002, table 7-6);
// before: both together were rejected and the extended position was switched off
IF ( ParCfg.Rob.OptionalCyclic.UseCartesianPositionExt AND NOT ParCfg.Rob.OptionalCyclic.UseCartesianPosition )
THEN
  // set to valid configuration
  ParCfg.Rob.OptionalCyclic.UseCartesianPosition    := TRUE;
 
  // Set info
  SetInfo( InfoID := RobotLibraryInfoIdEnum.INFO_RECV_EXT_CART_POS_NOT_USABLE_WITH_RECV_CART_POS, Overwrite := TRUE);
   
  // Create log entry
  CreateLogMessage( Timestamp   := SystemTime,
                    MessageType := MessageType.CMD,
                    Severity    := Severity.INFO,
                    MessageCode := 0,
                    MessageText := 'UseCartesianPositionExt cannot be used without UseCartesianPosition -> UseCartesianPosition is automatically activated');
END_IF


// Check configuration if optional cyclic JointPosition valid ?
// ST-FIX F137: the extended joint position cannot be used without the joint position -> the joint
// position is activated automatically (spec 6.4.2 and InfoID 16#6003, table 7-6); before: the check
// (both together rejected) was switched off with AND FALSE
IF ( ParCfg.Rob.OptionalCyclic.UseJointPositionExt AND NOT ParCfg.Rob.OptionalCyclic.UseJointPosition )
THEN
  // set to valid configuration
  ParCfg.Rob.OptionalCyclic.UseJointPosition    := TRUE;
 
  // Set info
  SetInfo( InfoID := RobotLibraryInfoIdEnum.INFO_RECV_EXT_JOINT_POS_NOT_USABLE_WITH_RECV_JOINT_POS, Overwrite := TRUE);
   
  // Create log entry
  CreateLogMessage( Timestamp   := SystemTime,
                    MessageType := MessageType.CMD,
                    Severity    := Severity.INFO,
                    MessageCode := 0,
                    MessageText := 'UseJointPositionExt cannot be used without UseJointPosition -> UseJointPosition is automatically activated');
END_IF
// EndRegion }}}

// Region ParCfg.Parameter.SynchronizationModes {{{

// Check ToolData synchronisation mode during startup
IF (( ParCfg.Plc.Parameter.SynchronizationModes.Tool[SyncTime.DURING_START_UP] <  SyncMode.NO_SYNCHRONIZATION ) OR
    ( ParCfg.Plc.Parameter.SynchronizationModes.Tool[SyncTime.DURING_START_UP] >= SyncMode.AUTOMATIC          )) // Automatic is not allowed during startup
THEN
  // ST-FIX F130: only the warning of the data set (spec: no error); the RobotTask is initialized,
  // the data set is not synchronized (SyncModesValid in the HandleSync... methods)
  SetWarning( WarningID := RobotLibraryWarningIdEnum.WARN_TOOL_DATA_SYNC_MODE_INVALID, Overwrite := TRUE );
   
  // Create log entry
  CreateLogMessagePara1 ( Timestamp   := SystemTime,
                          MessageType := MessageType.CMD,
                          Severity    := Severity.INFO,
                          MessageCode := 0,
                          MessageText :=                    'ParCfg.Plc.Parameter.SynchronizationModes.Tool[SyncTime.DURING_START_UP] invalid SyncMode {1}',
                          Para1       := SYNC_MODE_TO_STRING(ParCfg.Plc.Parameter.SynchronizationModes.Tool[SyncTime.DURING_START_UP]));
END_IF

// Check ToolData synchronisation mode after startup
IF (( ParCfg.Plc.Parameter.SynchronizationModes.Tool[SyncTime.AFTER_START_UP] < SyncMode.NO_SYNCHRONIZATION ) OR
    ( ParCfg.Plc.Parameter.SynchronizationModes.Tool[SyncTime.AFTER_START_UP] > SyncMode.AUTOMATIC          ))
THEN
  // ST-FIX F130: only the warning of the data set (spec: no error); the RobotTask is initialized,
  // the data set is not synchronized (SyncModesValid in the HandleSync... methods)
  SetWarning( WarningID := RobotLibraryWarningIdEnum.WARN_TOOL_DATA_SYNC_MODE_INVALID, Overwrite := TRUE);
   
  // Create log entry
  CreateLogMessagePara1 ( Timestamp   := SystemTime,
                          MessageType := MessageType.CMD,
                          Severity    := Severity.INFO,
                          MessageCode := 0,
                          MessageText :=                    'ParCfg.Plc.Parameter.SynchronizationModes.Tool[SyncTime.AFTER_START_UP] invalid SyncMode {1}',
                          Para1       := SYNC_MODE_TO_STRING(ParCfg.Plc.Parameter.SynchronizationModes.Tool[SyncTime.AFTER_START_UP]));
END_IF


// Check FrameData synchronisation mode during startup
IF (( ParCfg.Plc.Parameter.SynchronizationModes.Frame[SyncTime.DURING_START_UP] <  SyncMode.NO_SYNCHRONIZATION ) OR
    ( ParCfg.Plc.Parameter.SynchronizationModes.Frame[SyncTime.DURING_START_UP] >= SyncMode.AUTOMATIC          )) // Automatic is not allowed during startup
THEN
  // ST-FIX F130: only the warning of the data set (spec: no error); the RobotTask is initialized,
  // the data set is not synchronized (SyncModesValid in the HandleSync... methods)
  SetWarning( WarningID := RobotLibraryWarningIdEnum.WARN_FRAME_DATA_SYNC_MODE_INVALID, Overwrite := FALSE);
   
  // Create log entry
  CreateLogMessagePara1 ( Timestamp   := SystemTime,
                          MessageType := MessageType.CMD,
                          Severity    := Severity.INFO,
                          MessageCode := 0,
                          MessageText :=                    'ParCfg.Plc.Parameter.SynchronizationModes.Frame[SyncTime.DURING_START_UP] invalid SyncMode {1}',
                          Para1       := SYNC_MODE_TO_STRING(ParCfg.Plc.Parameter.SynchronizationModes.Frame[SyncTime.DURING_START_UP]));
END_IF


// Check FrameData synchronisation mode after startup
IF (( ParCfg.Plc.Parameter.SynchronizationModes.Frame[SyncTime.AFTER_START_UP] < SyncMode.NO_SYNCHRONIZATION ) OR
    ( ParCfg.Plc.Parameter.SynchronizationModes.Frame[SyncTime.AFTER_START_UP] > SyncMode.AUTOMATIC          ))
THEN
  // ST-FIX F130: only the warning of the data set (spec: no error); the RobotTask is initialized,
  // the data set is not synchronized (SyncModesValid in the HandleSync... methods)
  SetWarning( WarningID := RobotLibraryWarningIdEnum.WARN_FRAME_DATA_SYNC_MODE_INVALID, Overwrite := TRUE);
   
  // Create log entry
  CreateLogMessagePara1 ( Timestamp   := SystemTime,
                          MessageType := MessageType.CMD,
                          Severity    := Severity.INFO,
                          MessageCode := 0,
                          MessageText :=                    'ParCfg.Plc.Parameter.SynchronizationModes.Frame[SyncTime.AFTER_START_UP] invalid SyncMode {1}',
                          Para1       := SYNC_MODE_TO_STRING(ParCfg.Plc.Parameter.SynchronizationModes.Frame[SyncTime.AFTER_START_UP]));
END_IF


// Check LoadData synchronisation mode during startup
IF (( ParCfg.Plc.Parameter.SynchronizationModes.Load[SyncTime.DURING_START_UP] <  SyncMode.NO_SYNCHRONIZATION ) OR
    ( ParCfg.Plc.Parameter.SynchronizationModes.Load[SyncTime.DURING_START_UP] >= SyncMode.AUTOMATIC          )) // Automatic is not allowed during startup
THEN
  // ST-FIX F130: only the warning of the data set (spec: no error); the RobotTask is initialized,
  // the data set is not synchronized (SyncModesValid in the HandleSync... methods)
  SetWarning ( WarningID := RobotLibraryWarningIdEnum.WARN_LOAD_DATA_SYNC_MODE_INVALID, Overwrite := TRUE);
   
  // Create log entry
  CreateLogMessagePara1 ( Timestamp   := SystemTime,
                          MessageType := MessageType.CMD,
                          Severity    := Severity.INFO,
                          MessageCode := 0,
                          MessageText :=                    'ParCfg.Plc.Parameter.SynchronizationModes.Load[SyncTime.DURING_START_UP] invalid SyncMode {1}',
                          Para1       := SYNC_MODE_TO_STRING(ParCfg.Plc.Parameter.SynchronizationModes.Load[SyncTime.DURING_START_UP]));
END_IF


// Check LoadData synchronisation mode after startup
IF (( ParCfg.Plc.Parameter.SynchronizationModes.Load[SyncTime.AFTER_START_UP] < SyncMode.NO_SYNCHRONIZATION ) OR
    ( ParCfg.Plc.Parameter.SynchronizationModes.Load[SyncTime.AFTER_START_UP] > SyncMode.AUTOMATIC          ))
THEN
  // ST-FIX F130: only the warning of the data set (spec: no error); the RobotTask is initialized,
  // the data set is not synchronized (SyncModesValid in the HandleSync... methods)
  SetWarning( WarningID := RobotLibraryWarningIdEnum.WARN_LOAD_DATA_SYNC_MODE_INVALID, Overwrite := TRUE);
   
  // Create log entry
  CreateLogMessagePara1 ( Timestamp   := SystemTime,
                          MessageType := MessageType.CMD,
                          Severity    := Severity.INFO,
                          MessageCode := 0,
                          MessageText :=                    'ParCfg.Plc.Parameter.SynchronizationModes.Load[SyncTime.AFTER_START_UP] invalid SyncMode {1}',
                          Para1       := SYNC_MODE_TO_STRING(ParCfg.Plc.Parameter.SynchronizationModes.Load[SyncTime.AFTER_START_UP]));
END_IF


// Check WorkAreas synchronisation mode during startup
IF (( ParCfg.Plc.Parameter.SynchronizationModes.WorkAreas[SyncTime.DURING_START_UP] <  SyncMode.NO_SYNCHRONIZATION ) OR
    ( ParCfg.Plc.Parameter.SynchronizationModes.WorkAreas[SyncTime.DURING_START_UP] >= SyncMode.AUTOMATIC          )) // Automatic is not allowed during startup
THEN
  // ST-FIX F130: only the warning of the data set (spec: no error); the RobotTask is initialized,
  // the data set is not synchronized (SyncModesValid in the HandleSync... methods)
  SetWarning( WarningID := RobotLibraryWarningIdEnum.WARN_WORK_AREA_SYNC_MODE_INVALID, Overwrite := TRUE);
   
  // Create log entry
  CreateLogMessagePara1 ( Timestamp   := SystemTime,
                          MessageType := MessageType.CMD,
                          Severity    := Severity.INFO,
                          MessageCode := 0,
                          MessageText :=                    'ParCfg.Plc.Parameter.SynchronizationModes.WorkAreas[SyncTime.DURING_START_UP] invalid SyncMode {1}',
                          Para1       := SYNC_MODE_TO_STRING(ParCfg.Plc.Parameter.SynchronizationModes.WorkAreas[SyncTime.DURING_START_UP]));
END_IF


// Check WorkAreas synchronisation mode after startup
IF (( ParCfg.Plc.Parameter.SynchronizationModes.WorkAreas[SyncTime.AFTER_START_UP] < SyncMode.NO_SYNCHRONIZATION ) OR
    ( ParCfg.Plc.Parameter.SynchronizationModes.WorkAreas[SyncTime.AFTER_START_UP] > SyncMode.AUTOMATIC          ))
THEN
  // ST-FIX F130: only the warning of the data set (spec: no error); the RobotTask is initialized,
  // the data set is not synchronized (SyncModesValid in the HandleSync... methods)
  SetWarning( WarningID := RobotLibraryWarningIdEnum.WARN_WORK_AREA_SYNC_MODE_INVALID, Overwrite := TRUE);
   
  // Create log entry
  CreateLogMessagePara1 ( Timestamp   := SystemTime,
                          MessageType := MessageType.CMD,
                          Severity    := Severity.INFO,
                          MessageCode := 0,
                          MessageText :=                    'ParCfg.Plc.Parameter.SynchronizationModes.WorkAreas[SyncTime.AFTER_START_UP] invalid SyncMode {1}',
                          Para1       := SYNC_MODE_TO_STRING(ParCfg.Plc.Parameter.SynchronizationModes.WorkAreas[SyncTime.AFTER_START_UP]));
END_IF


// Check SWLimits synchronisation mode during startup
IF (( ParCfg.Plc.Parameter.SynchronizationModes.SWLimits[SyncTime.DURING_START_UP] <  SyncMode.NO_SYNCHRONIZATION ) OR
    ( ParCfg.Plc.Parameter.SynchronizationModes.SWLimits[SyncTime.DURING_START_UP] >= SyncMode.AUTOMATIC          )) // Automatic is not allowed during startup
THEN
  // ST-FIX F130: only the warning of the data set (spec: no error); the RobotTask is initialized,
  // the data set is not synchronized (SyncModesValid in the HandleSync... methods)
  SetWarning( WarningID := RobotLibraryWarningIdEnum.WARN_SW_LIMITS_SYNC_MODE_INVALID, Overwrite := TRUE);
   
  // Create log entry
  CreateLogMessagePara1 ( Timestamp   := SystemTime,
                          MessageType := MessageType.CMD,
                          Severity    := Severity.INFO,
                          MessageCode := 0,
                          MessageText :=                    'ParCfg.Plc.Parameter.SynchronizationModes.SWLimits[SyncTime.DURING_START_UP] invalid SyncMode {1}',
                          Para1       := SYNC_MODE_TO_STRING(ParCfg.Plc.Parameter.SynchronizationModes.SWLimits[SyncTime.DURING_START_UP]));
END_IF


// Check SWLimits synchronisation mode after startup
IF (( ParCfg.Plc.Parameter.SynchronizationModes.SWLimits[SyncTime.AFTER_START_UP] < SyncMode.NO_SYNCHRONIZATION ) OR
    ( ParCfg.Plc.Parameter.SynchronizationModes.SWLimits[SyncTime.AFTER_START_UP] > SyncMode.AUTOMATIC          ))
THEN
  // ST-FIX F130: only the warning of the data set (spec: no error); the RobotTask is initialized,
  // the data set is not synchronized (SyncModesValid in the HandleSync... methods)
  SetWarning( WarningID := RobotLibraryWarningIdEnum.WARN_SW_LIMITS_SYNC_MODE_INVALID, Overwrite := TRUE);
   
  // Create log entry
  CreateLogMessagePara1 ( Timestamp   := SystemTime,
                          MessageType := MessageType.CMD,
                          Severity    := Severity.INFO,
                          MessageCode := 0,
                          MessageText :=                    'ParCfg.Plc.Parameter.SynchronizationModes.SWLimits[SyncTime.AFTER_START_UP] invalid SyncMode {1}',
                          Para1       := SYNC_MODE_TO_STRING(ParCfg.Plc.Parameter.SynchronizationModes.SWLimits[SyncTime.AFTER_START_UP]));
END_IF


// Check DefaultDynamics synchronisation mode during startup
IF (( ParCfg.Plc.Parameter.SynchronizationModes.DefaultDynamics[SyncTime.DURING_START_UP] <  SyncMode.NO_SYNCHRONIZATION ) OR
    ( ParCfg.Plc.Parameter.SynchronizationModes.DefaultDynamics[SyncTime.DURING_START_UP] >= SyncMode.AUTOMATIC          )) // Automatic is not allowed during startup
THEN
  // ST-FIX F130: only the warning of the data set (spec: no error); the RobotTask is initialized,
  // the data set is not synchronized (SyncModesValid in the HandleSync... methods)
  SetWarning( WarningID := RobotLibraryWarningIdEnum.WARN_DEFAULT_DYNAMICS_SYNC_MODE_INVALID, Overwrite := TRUE);
   
  // Create log entry
  CreateLogMessagePara1 ( Timestamp   := SystemTime,
                          MessageType := MessageType.CMD,
                          Severity    := Severity.INFO,
                          MessageCode := 0,
                          MessageText :=                    'ParCfg.Plc.Parameter.SynchronizationModes.DefaultDynamics[SyncTime.DURING_START_UP] invalid SyncMode {1}',
                          Para1       := SYNC_MODE_TO_STRING(ParCfg.Plc.Parameter.SynchronizationModes.DefaultDynamics[SyncTime.DURING_START_UP]));
END_IF


// Check DefaultDynamics synchronisation mode after startup
IF (( ParCfg.Plc.Parameter.SynchronizationModes.DefaultDynamics[SyncTime.AFTER_START_UP] < SyncMode.NO_SYNCHRONIZATION ) OR
    ( ParCfg.Plc.Parameter.SynchronizationModes.DefaultDynamics[SyncTime.AFTER_START_UP] > SyncMode.AUTOMATIC          ))
THEN
  // ST-FIX F130: only the warning of the data set (spec: no error); the RobotTask is initialized,
  // the data set is not synchronized (SyncModesValid in the HandleSync... methods)
  SetWarning( WarningID := RobotLibraryWarningIdEnum.WARN_DEFAULT_DYNAMICS_SYNC_MODE_INVALID, Overwrite := TRUE);
   
  // Create log entry
  CreateLogMessagePara1 ( Timestamp   := SystemTime,
                          MessageType := MessageType.CMD,
                          Severity    := Severity.INFO,
                          MessageCode := 0,
                          MessageText :=                    'ParCfg.Plc.Parameter.SynchronizationModes.DefaultDynamics[SyncTime.AFTER_START_UP] invalid SyncMode {1}',
                          Para1       := SYNC_MODE_TO_STRING(ParCfg.Plc.Parameter.SynchronizationModes.DefaultDynamics[SyncTime.AFTER_START_UP]));
END_IF


// Check ReferenceDynamics synchronisation mode during startup
IF (( ParCfg.Plc.Parameter.SynchronizationModes.ReferenceDynamics[SyncTime.DURING_START_UP] <  SyncMode.NO_SYNCHRONIZATION ) OR
    ( ParCfg.Plc.Parameter.SynchronizationModes.ReferenceDynamics[SyncTime.DURING_START_UP] >= SyncMode.AUTOMATIC          )) // Automatic is not allowed during startup
THEN
  // ST-FIX F130: only the warning of the data set (spec: no error); the RobotTask is initialized,
  // the data set is not synchronized (SyncModesValid in the HandleSync... methods)
  SetWarning( WarningID := RobotLibraryWarningIdEnum.WARN_REFERENCE_DYNAMICS_SYNC_MODE_INVALID, Overwrite := TRUE);
   
  // Create log entry
  CreateLogMessagePara1 ( Timestamp   := SystemTime,
                          MessageType := MessageType.CMD,
                          Severity    := Severity.INFO,
                          MessageCode := 0,
                          MessageText :=                    'ParCfg.Plc.Parameter.SynchronizationModes.ReferenceDynamics[SyncTime.DURING_START_UP] invalid SyncMode {1}',
                          Para1       := SYNC_MODE_TO_STRING(ParCfg.Plc.Parameter.SynchronizationModes.ReferenceDynamics[SyncTime.DURING_START_UP]));
END_IF


// Check ReferenceDynamics synchronisation mode after startup
IF (( ParCfg.Plc.Parameter.SynchronizationModes.ReferenceDynamics[SyncTime.AFTER_START_UP] < SyncMode.NO_SYNCHRONIZATION ) OR
    ( ParCfg.Plc.Parameter.SynchronizationModes.ReferenceDynamics[SyncTime.AFTER_START_UP] > SyncMode.AUTOMATIC          ))
THEN
  // ST-FIX F130: only the warning of the data set (spec: no error); the RobotTask is initialized,
  // the data set is not synchronized (SyncModesValid in the HandleSync... methods)
  SetWarning( WarningID := RobotLibraryWarningIdEnum.WARN_REFERENCE_DYNAMICS_SYNC_MODE_INVALID, Overwrite := TRUE);
   
  // Create log entry
  CreateLogMessagePara1 ( Timestamp   := SystemTime,
                          MessageType := MessageType.CMD,
                          Severity    := Severity.INFO,
                          MessageCode := 0,
                          MessageText :=                    'ParCfg.Plc.Parameter.SynchronizationModes.ReferenceDynamics[SyncTime.AFTER_START_UP] invalid SyncMode {1}',
                          Para1       := SYNC_MODE_TO_STRING(ParCfg.Plc.Parameter.SynchronizationModes.ReferenceDynamics[SyncTime.AFTER_START_UP]));
END_IF
// EndRegion }}}
                
END_METHOD

METHOD PROTECTED CreateSendPayload : DINT
VAR_IN_OUT
  /// Robot assignment of function
  AxesGroup    : AxesGroup;
  /// Outputs of PLC for communication to RC
  RobotOutData : ARRAY[*] OF BYTE;
END_VAR
                  // ------------------------------------
// Fill SendData
// ------------------------------------
// Call SendData FB, update payload and size 
SendData( Payload := RobotOutData, PayLoadSize := ROBOT_OUT_DATA_SIZE);
// reset all variables and payload
SendData.Reset();

CreateSendPayloadHeader        ( AxesGroup := AxesGroup );
CreateSendPayloadCyclic        ( AxesGroup := AxesGroup );
CreateSendPayloadCyclicOptional( AxesGroup := AxesGroup );
CreateSendPayloadSequence      ( AxesGroup := AxesGroup );
CreateSendPayloadFooter        ( AxesGroup := AxesGroup );
CreateSendPayloadLogging       ( AxesGroup := AxesGroup );

// reset NewSEQ flag
AxesGroup.State.NewSEQ[0] := FALSE;
AxesGroup.State.NewSEQ[1] := FALSE; // ST-FIX F63: 2nd sequence was rebuilt in every cycle
                
END_METHOD

METHOD PROTECTED CreateSendPayloadCyclic : DINT
VAR_IN_OUT
  /// Robot assignment of function
  AxesGroup : AxesGroup;
END_VAR
                  // ST-FIX F2: ToolNo/FrameNo only with Cartesian Position RC -> PLC (spec table 5-88 bit 1)
IF ( AxesGroup.CyclicOptional.RobToPlc.CartesianPosition.Active )
THEN
  SendData.AddByte(Telegram.PlcToRob.Cyclic.ToolNo);
  SendData.AddByte(Telegram.PlcToRob.Cyclic.FrameNo);
END_IF

                
END_METHOD

METHOD PROTECTED CreateSendPayloadCyclicOptional : DINT
VAR_IN_OUT
  /// Robot assignment of function
  AxesGroup : AxesGroup;
END_VAR

VAR 
  /// temporary byte
 _tmpByte   : BYTE;
END_VAR
                  // Telegram.PlcToRob.CyclicOptional.SubProgramData {{{
IF ( AxesGroup.CyclicOptional.PlcToRob.SubProgramData.Active )
THEN
  SendData.AddDataBlock( ADR(Telegram.PlcToRob.CyclicOptional.SubProgramData.Data), SIZEOF(Telegram.PlcToRob.CyclicOptional.SubProgramData.Data));  
END_IF
// }}}
    
// Telegram.PlcToRob.CyclicOptional.CartesianPos {{{
IF ( AxesGroup.CyclicOptional.PlcToRob.CartesianPosition.Active) 
THEN
  SendData.AddReal(Telegram.PlcToRob.CyclicOptional.CartesianPosition.X );
  SendData.AddReal(Telegram.PlcToRob.CyclicOptional.CartesianPosition.Y );
  SendData.AddReal(Telegram.PlcToRob.CyclicOptional.CartesianPosition.Z );
  SendData.AddReal(Telegram.PlcToRob.CyclicOptional.CartesianPosition.Rx);
  SendData.AddReal(Telegram.PlcToRob.CyclicOptional.CartesianPosition.Ry);
  SendData.AddReal(Telegram.PlcToRob.CyclicOptional.CartesianPosition.Rz);

 _tmpByte   := 0;
 _tmpByte.0 := Telegram.PlcToRob.CyclicOptional.CartesianPosition.Config.0;
 _tmpByte.1 := Telegram.PlcToRob.CyclicOptional.CartesianPosition.Config.1;
 _tmpByte.2 := Telegram.PlcToRob.CyclicOptional.CartesianPosition.Config.2;
 
  SendData.AddByte(_tmpByte);
  SendData.AddByte(0); // ST-FIX F1: Config is 2 bytes (spec table 5-97)
          
  SendData.AddByte (Telegram.PlcToRob.CyclicOptional.CartesianPosition.Turns_J2_J1             );
  SendData.AddByte (Telegram.PlcToRob.CyclicOptional.CartesianPosition.Turns_J4_J3             );
  SendData.AddByte (Telegram.PlcToRob.CyclicOptional.CartesianPosition.Turns_J6_J5             );
  SendData.AddByte (Telegram.PlcToRob.CyclicOptional.CartesianPosition.Turns_E1                );
  SendData.AddReal (Telegram.PlcToRob.CyclicOptional.CartesianPosition.E1                      );
END_IF
// }}}

// Telegram.PlcToRob.CyclicOptional.JointPosition {{{
IF ( AxesGroup.CyclicOptional.PlcToRob.JointPosition.Active) 
THEN
  SendData.AddReal(Telegram.PlcToRob.CyclicOptional.JointPosition.J1);
  SendData.AddReal(Telegram.PlcToRob.CyclicOptional.JointPosition.J2);
  SendData.AddReal(Telegram.PlcToRob.CyclicOptional.JointPosition.J3);
  SendData.AddReal(Telegram.PlcToRob.CyclicOptional.JointPosition.J4);
  SendData.AddReal(Telegram.PlcToRob.CyclicOptional.JointPosition.J5);
  SendData.AddReal(Telegram.PlcToRob.CyclicOptional.JointPosition.J6);
  SendData.AddReal(Telegram.PlcToRob.CyclicOptional.JointPosition.E1);
END_IF
// }}}

// Telegram.PlcToRob.CyclicOptional.Force {{{
IF ( AxesGroup.CyclicOptional.PlcToRob.Force.Active) 
THEN
  SendData.AddReal(Telegram.PlcToRob.CyclicOptional.Force.X);
  SendData.AddReal(Telegram.PlcToRob.CyclicOptional.Force.Y);
  SendData.AddReal(Telegram.PlcToRob.CyclicOptional.Force.Z);
  SendData.AddReal(Telegram.PlcToRob.CyclicOptional.Force.Rx);
  SendData.AddReal(Telegram.PlcToRob.CyclicOptional.Force.Ry);
  SendData.AddReal(Telegram.PlcToRob.CyclicOptional.Force.Rz);
END_IF  
// }}}

// Telegram.PlcToRob.CyclicOptional.TwoSequences {{{
// }}}

// AxesGroup.OptionalCyclic.PlcToRob.CartesianPosExt {{{
IF ( AxesGroup.CyclicOptional.PlcToRob.CartesianPositionExt.Active) 
THEN
  SendData.AddReal(Telegram.PlcToRob.CyclicOptional.CartesianPositionExt.E2);
  SendData.AddReal(Telegram.PlcToRob.CyclicOptional.CartesianPositionExt.E3);
  SendData.AddReal(Telegram.PlcToRob.CyclicOptional.CartesianPositionExt.E4);
  SendData.AddReal(Telegram.PlcToRob.CyclicOptional.CartesianPositionExt.E5);
  SendData.AddReal(Telegram.PlcToRob.CyclicOptional.CartesianPositionExt.E6);
END_IF    
// }}}

// AxesGroup.OptionalCyclic.PlcToRob.JointPositionExt {{{
IF ( AxesGroup.CyclicOptional.PlcToRob.JointPositionExt.Active) 
THEN
  SendData.AddReal(Telegram.PlcToRob.CyclicOptional.JointPositionExt.E2);
  SendData.AddReal(Telegram.PlcToRob.CyclicOptional.JointPositionExt.E3);  
  SendData.AddReal(Telegram.PlcToRob.CyclicOptional.JointPositionExt.E4);
  SendData.AddReal(Telegram.PlcToRob.CyclicOptional.JointPositionExt.E5);
  SendData.AddReal(Telegram.PlcToRob.CyclicOptional.JointPositionExt.E6);        
END_IF  
// }}}
                    
// Telegram.PlcToRob.CyclicOptional..CartesianForceExt {{{
IF ( AxesGroup.CyclicOptional.PlcToRob.ForceExt.Active) 
THEN
  SendData.AddReal(Telegram.PlcToRob.CyclicOptional.ForceExt.E1);
  SendData.AddReal(Telegram.PlcToRob.CyclicOptional.ForceExt.E2);
  SendData.AddReal(Telegram.PlcToRob.CyclicOptional.ForceExt.E3);
  SendData.AddReal(Telegram.PlcToRob.CyclicOptional.ForceExt.E4);
  SendData.AddReal(Telegram.PlcToRob.CyclicOptional.ForceExt.E5);
  SendData.AddReal(Telegram.PlcToRob.CyclicOptional.ForceExt.E6);
END_IF                    
// }}}
                
END_METHOD

METHOD PRIVATE CreateSendPayloadFooter : DINT
VAR_IN_OUT
  /// Robot assignment of function
  AxesGroup : AxesGroup;
END_VAR
VAR
END_VAR
                  SendData.SetLifeSignFooter( LifeSign :=  AxesGroup.Cyclic.PlcToRob.LifeSign);

                
END_METHOD

METHOD PROTECTED CreateSendPayloadHeader : DINT
VAR_IN_OUT
  /// Robot assignment of function
  AxesGroup : AxesGroup;
END_VAR
                  SendData.AddByte(Telegram.PlcToRob.Header.SRCIVersion           );
SendData.AddByte(Telegram.PlcToRob.Header.FastStop_LifeSign     ); 
SendData.AddUint(Telegram.PlcToRob.Header.TelegramLengthPlcToRob);
SendData.AddUint(Telegram.PlcToRob.Header.TelegramLengthRobToPlc);
SendData.AddByte(Telegram.PlcToRob.Header.AxesGroupID_Control   );
SendData.AddByte(Telegram.PlcToRob.Header.Reserved              );
SendData.AddUint(Telegram.PlcToRob.Header.TelegramNumberPlcToRob);
SendData.AddUint(Telegram.PlcToRob.Header.TelegramNumberRobToPlc);
SendData.AddUint(Telegram.PlcToRob.Header.ClientDate            ); 
SendData.AddTime(Telegram.PlcToRob.Header.ClientTime            );  
                
END_METHOD

METHOD PRIVATE CreateSendPayloadLogging : DINT
VAR_IN_OUT
  /// Robot assignment of function
  AxesGroup                 : AxesGroup;
END_VAR
                  IF  ((( Telegram.PlcToRob.Sequence[0].Header.PayloadLength > 0 ) AND (AxesGroup.State.NewSEQ[0] )) OR
     (( Telegram.PlcToRob.Sequence[1].Header.PayloadLength > 0 ) AND (AxesGroup.State.NewSEQ[1] )))
THEN
  // Create log entry
  CreateLogMessagePara1 ( Timestamp   := SystemTime,
                          MessageType := MessageType.CMD,
                          Severity    := Severity.DEBUG,
                          MessageCode := 0,
                          MessageText := 'SendData: Bytes send in total: {1}',
                          Para1       :=  UDINT_TO_STRING(SendData.PayloadLen));
END_IF
                
END_METHOD

METHOD PRIVATE CreateSendPayloadSequence : DINT
VAR_IN_OUT
  /// Robot assignment of function
  AxesGroup                 : AxesGroup;
END_VAR

VAR 
  /// internal sequence index
 _seqIdx                    : DINT;
  /// internal fragment index
 _fragIdx                   : DINT;
END_VAR
                  FOR _seqIdx := 0 TO AxesGroup.State.SequenceCountSend
DO
  // ST-FIX F63: every telegram sequence starts at its own address (Fig. 5-205); before, the
  // 1st sequence ran into the area of the 2nd one and the 2nd header was sent only sometimes
  IF ( _seqIdx = PRIMARY_SEQUENCE )
  THEN
    SendData.PayloadPtr := CalculateSequencePayloadStartAdr(AxesGroup := AxesGroup, 
                                                            Direction := ComDirection.PLC_TO_ROB,
                                                            Sequence  := SequenceFlag.PRIMARY_SEQUENCE);
  ELSE
    SendData.PayloadPtr := CalculateSequencePayloadStartAdr(AxesGroup := AxesGroup, 
                                                            Direction := ComDirection.PLC_TO_ROB,
                                                            Sequence  := SequenceFlag.SECONDARY_SEQUENCE);
  END_IF

  // Telegram.PlcToRob.Sequence[x].Header {{{
  SendData.AddUint(Telegram.PlcToRob.Sequence[_seqIdx].Header.SEQ_ACK);
  SendData.AddUint(Telegram.PlcToRob.Sequence[_seqIdx].Header.PayloadLength);
  // }}}

  // check limit reachted ?
  IF ( SendData.PayloadPtr + FOOTER_SIZE >= Telegram.PlcToRob.Header.TelegramLengthPlcToRob)
  THEN
    EXIT;
  END_IF
  
  // PlcToRob.Sequence[x].Fragment[x] {{{
  FOR _fragIdx := 0 TO AxesGroup.State.FragmentCountSend[_seqIdx]  
  DO

    IF (Telegram.PlcToRob.Sequence[_seqIdx].Fragment[_fragIdx].Header.PayloadLength > 0)
    THEN  
      // PlcToRob.Sequence[x].Fragment[x].Header {{{        
      SendData.AddUint(Telegram.PlcToRob.Sequence[_seqIdx].Fragment[_fragIdx].Header.CmdID);
      SendData.AddByte(Telegram.PlcToRob.Sequence[_seqIdx].Fragment[_fragIdx].Header.Reserve);
      SendData.AddByte(Telegram.PlcToRob.Sequence[_seqIdx].Fragment[_fragIdx].Header.FragmentAction);
      SendData.AddUint(Telegram.PlcToRob.Sequence[_seqIdx].Fragment[_fragIdx].Header.PayloadPointer);
      SendData.AddUint(Telegram.PlcToRob.Sequence[_seqIdx].Fragment[_fragIdx].Header.PayloadLength);
      // }}}
      
      // PlcToRob.Sequence[x].Fragment[x].Command {{{
      
      // Hint: the command header is part of the fragment payload  
      IF (Telegram.PlcToRob.Sequence[_seqIdx].Fragment[_fragIdx].Header.PayloadLength > 0)
      THEN
        SendData.AddDataBlock( pValue :=  ADR(Telegram.PlcToRob.Sequence[_seqIdx].Fragment[_fragIdx].Command.Payload           ) + Telegram.PlcToRob.Sequence[_seqIdx].Fragment[_fragIdx].Header.PayloadPointer,
                                 Size :=     (Telegram.PlcToRob.Sequence[_seqIdx].Fragment[_fragIdx].Header.PayloadLength      ));

      END_IF
      
      
      IF (SendData.PayloadLen = 232)
      THEN
        SendData.PayloadLen := SendData.PayloadLen;
			END_IF
      
    END_IF
    // }}}
  END_FOR
  // }}}
END_FOR  
                
END_METHOD

METHOD FB_init : BOOL
VAR_INPUT
  bInitRetains : BOOL; // if TRUE, the retain variables are initialized (warm start / cold start)
  bInCopyCode : BOOL;  // if TRUE, the instance afterwards gets moved into the copy code (online change)
END_VAR
                  MyType := 'MC_RobotTaskFB';

// ST-FIX F132: identification of this instance (an online change keeps the old value)
IF ( NOT bInCopyCode )
THEN
 _instanceCount := _instanceCount + 1;
 _instanceId    := _instanceCount;
END_IF

// Create log entry
CreateLogMessage ( Timestamp   := SystemTime,
                   MessageType := MessageType.CMD,
                   Severity    := Severity.DEBUG,
                   MessageCode := 0,
                   MessageText := 'PLC started / restarted');

                
END_METHOD

METHOD PRIVATE HandleAliveBit
VAR_INPUT
  LifeSign : BYTE;
END_VAR

VAR_INST
  /// flag that indicates that the 1st cyclce is running
  First : BOOL := TRUE;
END_VAR
                  IF (First AND LifeSign > 0)
THEN
  // init alive value
 _aliveValue := LifeSign;
  // reset first flag
  First := FALSE;
END_IF

_aliveCheck ( IN  := Enable AND (_aliveValue = LifeSign) (* ST-FIX F181: only while enabled *), PT := ParCfg.Com.LifeSignTimeOut + ParCfg.Plc.CycleTime);
_alive_R    ( CLK := _aliveBit);
_alive_F    ( CLK := _aliveBit);

IF ( _aliveValue <> LifeSign)
THEN
 _aliveValue := LifeSign;
 _aliveBit   := TRUE;
END_IF

IF (_aliveCheck.Q)
THEN
 _aliveBit := FALSE;
END_IF

IF (_alive_R.Q)
THEN
  // Create log entry
  CreateLogMessage ( Timestamp   := SystemTime,
                     MessageType := MessageType.CMD,
                     Severity    := Severity.INFO,
                     MessageCode := 0,
                     MessageText := 'Data Exchange is running (Alive-Bit)');
END_IF

IF (_alive_F.Q)
THEN
  // Create log entry
  CreateLogMessage ( Timestamp   := SystemTime,
                     MessageType := MessageType.CMD,
                     Severity    := Severity.INFO,
                     MessageCode := 0,
                     MessageText := 'Data Exchange has stopped (Alive-Bit)');
END_IF

                
END_METHOD

METHOD PRIVATE HandleAxesGroup
VAR_IN_OUT
  /// Robot assignment of function
  AxesGroup         : AxesGroup;
  /// ToolData stored on PLC. For more information refer to 5.5.6.3
  ToolData          : ARRAY[*] OF Tool;
  /// LoadData stored on PLC.For more information refer to 5.5.6.4
  FrameData         : ARRAY[*] OF Frame;
  /// LoadData stored on PLC.For more information refer to 5.5.6.4 
  LoadData          : ARRAY[*] OF Load;
  /// Work areas stored on PLC. For more information refer to 5.5.8
  WorkAreas         : ARRAY[*] OF RobotWorkArea;
  /// Software limits stored on PLC
  SWLimits          : SWLimits;
  /// Default dynamics stored on PLC. For more information refer to 5.5.7
  DefaultDynamics   : DefaultDynamics;
  /// Reference dynamics stored on PLC. For more information refer to 5.5.7
  ReferenceDynamics : ReferenceDynamics;  
END_VAR
                  HandleAxesGroupAcyclic       ( AxesGroup         := AxesGroup );
HandleAxesGroupCyclic        ( AxesGroup         := AxesGroup );
HandleAxesGroupCyclicOptional( AxesGroup         := AxesGroup );
HandleAxesGroupMessageLog    ( AxesGroup         := AxesGroup );
HandleAxesGroupParameter     ( AxesGroup         := AxesGroup );
HandleAxesGroupState         ( AxesGroup         := AxesGroup );
HandleAxesGroupSystemData    ( AxesGroup         := AxesGroup, 
	                             ToolData          := ToolData, 
	                             FrameData         := FrameData, 
	                             LoadData          := LoadData, 
	                             WorkAreas         := WorkAreas, 
	                             SWLimits          := SWLimits, 
	                             DefaultDynamics   := DefaultDynamics, 
	                             ReferenceDynamics := ReferenceDynamics);
                
END_METHOD

METHOD PRIVATE HandleAxesGroupAcyclic
VAR_IN_OUT
  /// Robot assignment of function
  AxesGroup : AxesGroup;
END_VAR
                  // Call active command register FB
AxesGroup.Acyclic.ActiveCommandRegister(SystemTime     := SystemTime,
                                        RegisterSize   := MIN( RobotLibraryParameter.ACTIVE_CMD_REGISTER_ENTRIES_MAX, AxesGroup.Parameter.Rob.Parameter.LengthACR),
                                        InternalLogger := AxesGroup.MessageLog, 
                                        ExternalLogger := AxesGroup.MessageLog.ExternalLogger,
                                        LogLevel       := AxesGroup.MessageLog.LogLevel);
                
END_METHOD

METHOD PRIVATE HandleAxesGroupCyclic
VAR_IN_OUT
  /// Robot assignment of function
  AxesGroup : AxesGroup;
END_VAR
                  // set instance AxesGroupID
AxesGroup.Cyclic.PlcToRob.AxesGroupID := AxesGroupID;
// Set Version
AxesGroup.Cyclic.PlcToRob.SRCIVersion := RobotLibraryConstants.SRCIVersion;

AxesGroup.Cyclic.PlcToRob.TelegramLengthPlcToRob := _parCfg.Com.TelegramLengthPlcToRob;
AxesGroup.Cyclic.PlcToRob.TelegramLengthRobToPlc := _parCfg.Com.TelegramLengthRobToPlc;

AxesGroup.Cyclic.PlcToRob.TelegramNumberPlcToRob := PlcOptionalCyclicToUint(AxesGroup.Parameter.Plc.OptionalCyclic);
AxesGroup.Cyclic.PlcToRob.TelegramNumberRobToPlc := RobOptionalCyclicToUint(AxesGroup.Parameter.Rob.OptionalCyclic);

// Set Date + Time
AxesGroup.Cyclic.PlcToRob.ClientDate  := DATE_TO_IEC_DATE(SystemTime.SystemDate);
AxesGroup.Cyclic.PlcToRob.ClientTime  := TIME_TO_IEC_TIME(SystemTime.SystemTime);
                
END_METHOD

METHOD PRIVATE HandleAxesGroupCyclicOptional
VAR_IN_OUT
  /// Robot assignment of function
  AxesGroup : AxesGroup;
END_VAR
                  // PlcToRob {{{
AxesGroup.CyclicOptional.PlcToRob.SubProgramData      .Active := AxesGroup.Parameter.Plc.OptionalCyclic.UseCallSubprogram; 
AxesGroup.CyclicOptional.PlcToRob.CartesianPosition   .Active := AxesGroup.Parameter.Plc.OptionalCyclic.UseCartesianPosition; 
AxesGroup.CyclicOptional.PlcToRob.JointPosition       .Active := AxesGroup.Parameter.Plc.OptionalCyclic.UseJointPosition; 
AxesGroup.CyclicOptional.PlcToRob.Force               .Active := AxesGroup.Parameter.Plc.OptionalCyclic.UseForce; 
AxesGroup.CyclicOptional.PlcToRob.CartesianPositionExt.Active := AxesGroup.Parameter.Plc.OptionalCyclic.UseCartesianPositionExt; 
AxesGroup.CyclicOptional.PlcToRob.JointPositionExt    .Active := AxesGroup.Parameter.Plc.OptionalCyclic.UseJointPositionExt; 
// }}}

// RobToPlc {{{
AxesGroup.CyclicOptional.RobToPlc.SubProgramData      .Active := AxesGroup.Parameter.Rob.OptionalCyclic.UseCallSubprogram; 
AxesGroup.CyclicOptional.RobToPlc.CartesianPosition   .Active := AxesGroup.Parameter.Rob.OptionalCyclic.UseCartesianPosition;    
AxesGroup.CyclicOptional.RobToPlc.JointPosition       .Active := AxesGroup.Parameter.Rob.OptionalCyclic.UseJointPosition;    
AxesGroup.CyclicOptional.RobToPlc.Force               .Active := AxesGroup.Parameter.Rob.OptionalCyclic.UseForce;
AxesGroup.CyclicOptional.RobToPlc.Current             .Active := AxesGroup.Parameter.Rob.OptionalCyclic.UseCurrent;    
AxesGroup.CyclicOptional.RobToPlc.CartesianPositionExt.Active := AxesGroup.Parameter.Rob.OptionalCyclic.UseCartesianPositionExt;    
AxesGroup.CyclicOptional.RobToPlc.JointPositionExt    .Active := AxesGroup.Parameter.Rob.OptionalCyclic.UseJointPositionExt;    
AxesGroup.CyclicOptional.RobToPlc.ForceExt            .Active := AxesGroup.Parameter.Rob.OptionalCyclic.UseForceExt;    
AxesGroup.CyclicOptional.RobToPlc.CurrentExt          .Active := AxesGroup.Parameter.Rob.OptionalCyclic.UseCurrentExt;    
// }}}

                
END_METHOD

METHOD PRIVATE HandleAxesGroupMessageLog
VAR_IN_OUT
  /// Robot assignment of function
  AxesGroup  : AxesGroup;
END_VAR
                  // Set External logger 
AxesGroup.MessageLog.ExternalLogger := ExternalLogger;
AxesGroup.MessageLog.LogLevel       := LogLevel;


IF (AxesGroup.State.GroupReset_R.Q)
THEN
  AxesGroup.MessageLog.DeleteMessages();
  AxesGroup.MessageLog.DeleteSystemLogs();
END_IF
                
END_METHOD

METHOD PRIVATE HandleAxesGroupParameter
VAR_IN_OUT
  /// Robot assignment of function
  AxesGroup : AxesGroup;
END_VAR
                  IF (_exchangeConfiguration.Enabled)
THEN
  AxesGroup.Parameter.Plc.Parameter                           := _parCfg.Plc.Parameter;      
  AxesGroup.Parameter.Plc.OptionalCyclic                      := _parCfg.Plc.OptionalCyclic;
  AxesGroup.Parameter.Rob.OptionalCyclic                      := _parCfg.Rob.OptionalCyclic;
  
  AxesGroup.Parameter.Rob.Parameter.LengthACR                 := _exchangeConfiguration.OutCmd.LengthACR;
  AxesGroup.Parameter.Rob.Parameter.HighestToolIndex          := _exchangeConfiguration.OutCmd.HighestToolIndex;
  AxesGroup.Parameter.Rob.Parameter.HighestFrameIndex         := _exchangeConfiguration.OutCmd.HighestFrameIndex;
  AxesGroup.Parameter.Rob.Parameter.HighestLoadIndex          := _exchangeConfiguration.OutCmd.HighestLoadIndex;
  AxesGroup.Parameter.Rob.Parameter.HighestWorkAreaIndex      := _exchangeConfiguration.OutCmd.HighestWorkAreaIndex;
  AxesGroup.Parameter.Rob.Parameter.DataInSync                := _exchangeConfiguration.OutCmd.DataInSync;
  AxesGroup.Parameter.Rob.Parameter.ChangeIndexTool           := _exchangeConfiguration.OutCmd.ChangeIndexTool;
  AxesGroup.Parameter.Rob.Parameter.ChangeIndexFrame          := _exchangeConfiguration.OutCmd.ChangeIndexFrame;
  AxesGroup.Parameter.Rob.Parameter.ChangeIndexLoad           := _exchangeConfiguration.OutCmd.ChangeIndexLoad;
  AxesGroup.Parameter.Rob.Parameter.ChangeIndexWorkArea       := _exchangeConfiguration.OutCmd.ChangeIndexWorkArea;
  AxesGroup.Parameter.Rob.Parameter.RAWorkingHours            := _exchangeConfiguration.OutCmd.RAWorkingHours;
  AxesGroup.Parameter.Rob.Parameter.BrakeTestRequired         := _exchangeConfiguration.OutCmd.BrakeTestRequired;
  AxesGroup.Parameter.Rob.Parameter.StepModeExactStopActive   := _exchangeConfiguration.OutCmd.StepModeExactStopActive;
  AxesGroup.Parameter.Rob.Parameter.StepModeBlendingActive    := _exchangeConfiguration.OutCmd.StepModeBlendingActive;
  AxesGroup.Parameter.Rob.Parameter.PathAccuracyMode          := _exchangeConfiguration.OutCmd.PathAccuracyMode;
  AxesGroup.Parameter.Rob.Parameter.AvoidSingularity          := _exchangeConfiguration.OutCmd.AvoidSingularity;
  AxesGroup.Parameter.Rob.Parameter.CollisionDetectionEnabled := _exchangeConfiguration.OutCmd.CollisionDetectionEnabled;
  AxesGroup.Parameter.Rob.Parameter.AcceleratingSupported     := _exchangeConfiguration.OutCmd.AcceleratingSupported;
  AxesGroup.Parameter.Rob.Parameter.DecceleratingSupported    := _exchangeConfiguration.OutCmd.DecceleratingSupported;
  AxesGroup.Parameter.Rob.Parameter.ConstantVelocitySupported := _exchangeConfiguration.OutCmd.ConstantVelocitySupported;
  AxesGroup.Parameter.Rob.Parameter.RCWorkingHours            := _exchangeConfiguration.OutCmd.RCWorkingHours;
ELSIF ( _stepCmd > 0 )
THEN
  // ST-FIX F151: while the RobotTask initializes, use the configuration taken at the enable
  // (_parCfg, including the corrections of CheckParameterValid, e.g. F137); the input ParCfg is
  // written again by the caller in every cycle and would change the telegram number during the start-up
  AxesGroup.Parameter.Plc.Parameter                           := _parCfg.Plc.Parameter;
  AxesGroup.Parameter.Plc.OptionalCyclic                      := _parCfg.Plc.OptionalCyclic;
  AxesGroup.Parameter.Rob.OptionalCyclic                      := _parCfg.Rob.OptionalCyclic;
ELSE
  AxesGroup.Parameter.Plc.Parameter                           := ParCfg.Plc.Parameter;      
  AxesGroup.Parameter.Plc.OptionalCyclic                      := ParCfg.Plc.OptionalCyclic;
  AxesGroup.Parameter.Rob.OptionalCyclic                      := ParCfg.Rob.OptionalCyclic;
END_IF
                
END_METHOD

METHOD PRIVATE HandleAxesGroupState
VAR_IN_OUT
  /// Robot assignment of function
  AxesGroup : AxesGroup;
END_VAR
VAR
  /// internal index for loops
 _idx       : DINT; 
END_VAR
                  AxesGroup.State.AliveOk      := _aliveBit;
AxesGroup.State.Initialized  := Initialized  AND AxesGroup.State.AliveOk;
AxesGroup.State.Synchronized := Synchronized AND AxesGroup.State.AliveOk;
AxesGroup.State.CMDsEnabled  := AxesGroup.State.Initialized OR 
                                AxesGroup.State.Synchronized;

AxesGroup.State.StatusRobotArm  := AxesGroup.Cyclic.RobToPlc.StatusRobotArm;                                
AxesGroup.State.ConfigExchanged := _exchangeConfiguration.Enabled;

AxesGroup.State.UnifiedFrameIndex                    := DINT_TO_USINT( MIN( MIN(AxesGroup.SystemData.FrameDataMax, RobotLibraryParameter.FRAME_MAX - 1), _exchangeConfiguration.OutCmd.HighestFrameIndex   ));
AxesGroup.State.UnifiedToolIndex                     := DINT_TO_USINT( MIN( MIN(AxesGroup.SystemData.ToolDataMax , RobotLibraryParameter.TOOL_MAX - 1), _exchangeConfiguration.OutCmd.HighestToolIndex    ));
AxesGroup.State.UnifiedLoadIndex                     := DINT_TO_USINT( MIN( MIN(AxesGroup.SystemData.LoadDataMax , RobotLibraryParameter.LOAD_MAX - 1), _exchangeConfiguration.OutCmd.HighestLoadIndex    ));
AxesGroup.State.UnifiedWorkAreaIndex                 := DINT_TO_USINT( MIN( MIN(AxesGroup.SystemData.WorkAreasMax, RobotLibraryParameter.WORK_AREAS_MAX - 1), _exchangeConfiguration.OutCmd.HighestWorkAreaIndex));

AxesGroup.State.DataEnableSync                       := _exchangeConfiguration.ParCmd.DataEnableSync;
AxesGroup.State.SyncStateRc.InSync.Frame             := _exchangeConfiguration.OutCmd.DataInSync.FramesInSync;
AxesGroup.State.SyncStateRc.InSync.Tool              := _exchangeConfiguration.OutCmd.DataInSync.ToolsInSync;
AxesGroup.State.SyncStateRc.InSync.Load              := _exchangeConfiguration.OutCmd.DataInSync.LoadsInSync;
AxesGroup.State.SyncStateRc.InSync.WorkArea          := _exchangeConfiguration.OutCmd.DataInSync.WorkAreasInSync;
AxesGroup.State.SyncStateRc.InSync.SwLimits          := _exchangeConfiguration.OutCmd.DataInSync.SoftwareLimitsInSync;
AxesGroup.State.SyncStateRc.InSync.DefaultDynamics   := _exchangeConfiguration.OutCmd.DataInSync.DefaultDynamicsInSync;
AxesGroup.State.SyncStateRc.InSync.ReferenceDynamics := _exchangeConfiguration.OutCmd.DataInSync.ReferenceDynamicsInSync;

AxesGroup.State.SyncStateRc.UnSyncNo.Frame           := _exchangeConfiguration.OutCmd.ChangeIndexFrame;
AxesGroup.State.SyncStateRc.UnSyncNo.Tool            := _exchangeConfiguration.OutCmd.ChangeIndexTool;
AxesGroup.State.SyncStateRc.UnSyncNo.Load            := _exchangeConfiguration.OutCmd.ChangeIndexLoad;
AxesGroup.State.SyncStateRc.UnSyncNo.WorkArea        := _exchangeConfiguration.OutCmd.ChangeIndexWorkArea;

// Update internal data
AxesGroup.State.SystemTime   := SystemTime;
AxesGroup.State.OnlineChange := OnlineChange;
AxesGroup.State.Initialized  := Initialized;

// Create rising and falling edges for Online Change
AxesGroup.State.OnlineChange_R(CLK := OnlineChange);
AxesGroup.State.OnlineChange_F(CLK := OnlineChange);

// Create rising and falling edges for GroupReset
AxesGroup.State.GroupReset_R(CLK := AxesGroup.State.GroupReset);
AxesGroup.State.GroupReset_F(CLK := AxesGroup.State.GroupReset);

// Copy function block results 
AxesGroup.State.RobotData         := _readRobotData.OutCmd;
AxesGroup.State.ConfigurationData := _exchangeConfiguration.OutCmd;
                
                
END_METHOD

METHOD PRIVATE HandleAxesGroupSystemData
VAR_IN_OUT
  /// Robot assignment of function
  AxesGroup         : AxesGroup;
  /// ToolData stored on PLC. For more information refer to 5.5.6.3
  ToolData          : ARRAY[*] OF Tool;
  /// LoadData stored on PLC.For more information refer to 5.5.6.4
  FrameData         : ARRAY[*] OF Frame;
  /// LoadData stored on PLC.For more information refer to 5.5.6.4 
  LoadData          : ARRAY[*] OF Load;
  /// Work areas stored on PLC. For more information refer to 5.5.8
  WorkAreas         : ARRAY[*] OF RobotWorkArea;
  /// Software limits stored on PLC
  SWLimits          : SWLimits;
  /// Default dynamics stored on PLC. For more information refer to 5.5.7
  DefaultDynamics   : DefaultDynamics;
  /// Reference dynamics stored on PLC. For more information refer to 5.5.7
  ReferenceDynamics : ReferenceDynamics;  
END_VAR
                  // Update ToolData                    
AxesGroup.SystemData.ToolDataPtr       := ToolData;
AxesGroup.SystemData.ToolDataMin       := LOWER_BOUND  (ToolData,1);
AxesGroup.SystemData.ToolDataMax       := UPPER_BOUND  (ToolData,1);
AxesGroup.SystemData.ToolDataCount     := DINT_TO_UDINT(1 + AxesGroup.SystemData.ToolDataMax - AxesGroup.SystemData.ToolDataMin);
                                       
// Update LoadData                    
AxesGroup.SystemData.LoadDataPtr       := LoadData;
AxesGroup.SystemData.LoadDataMin       := LOWER_BOUND  (LoadData,1);                                                    
AxesGroup.SystemData.LoadDataMax       := UPPER_BOUND  (LoadData,1);                                                    
AxesGroup.SystemData.LoadDataCount     := DINT_TO_UDINT(1 + AxesGroup.SystemData.LoadDataMax - AxesGroup.SystemData.LoadDataMin);
                                       
// Update FrameData       
AxesGroup.SystemData.FrameDataPtr      := FrameData;                                                                       
AxesGroup.SystemData.FrameDataMin      := LOWER_BOUND  (FrameData,1);                                                     
AxesGroup.SystemData.FrameDataMax      := UPPER_BOUND  (FrameData,1);                                                     
AxesGroup.SystemData.FrameDataCount    := DINT_TO_UDINT(1 + AxesGroup.SystemData.FrameDataMax - AxesGroup.SystemData.FrameDataMin);

// Update WorkAreas 
AxesGroup.SystemData.WorkAreasPtr      := WorkAreas;                                                                      
AxesGroup.SystemData.WorkAreasMin      := LOWER_BOUND  (WorkAreas,1);                                                     
AxesGroup.SystemData.WorkAreasMax      := UPPER_BOUND  (WorkAreas,1);                                                     
AxesGroup.SystemData.WorkAreasCount    := DINT_TO_UDINT(1 + AxesGroup.SystemData.WorkAreasMax - AxesGroup.SystemData.WorkAreasMin);

// Update SoftwareLimits 
AxesGroup.SystemData.SWLimits          REF= SWLimits;
// Update DefaultDynamics 
AxesGroup.SystemData.DefaultDynamics   REF= DefaultDynamics;
// Update ReferenceDynamics 
AxesGroup.SystemData.ReferenceDynamics REF= ReferenceDynamics;
                
                
END_METHOD

METHOD PRIVATE HandleInvalidFrames
VAR_IN_OUT
   /// Robot assignment of function
  AxesGroup   : AxesGroup;
    /// Inputs of PLC for communication from RC
  RobotInData : ARRAY[*] OF BYTE;
END_VAR 
VAR
  /// Value of lifesign in header
 _lifeSignHeader    : BYTE;
  /// Value of lifesign in footer
 _lifeSignFooter    : BYTE;
END_VAR
VAR_INST
  /// Timeout for invalid frames counter check
 _invalidFrameCounterCheck_D : TON;
  /// last count of invalid frames
 _lastInvalidFrames          : UDINT;
END_VAR
                  IF ( AxesGroup.Cyclic.RobToPlc.TelegramState = TelegramState.INITIALIZED ) 
THEN
  // Get lifesign values
 _lifeSignHeader := GetHalfeByteHi( RobotInData[ROBOT_IN_DATA_MIN + 1]);
 _lifeSignFooter := GetHalfeByteHi( RobotInData[MIN(ROBOT_IN_DATA_MIN + _parCfg.Com.TelegramLengthRobToPlc - 1,
                                                     ROBOT_IN_DATA_MAX)]); // ST-FIX F66: last byte of the telegram
END_IF

// Timer for invalid frame(s) message
_invalidFrameCounterCheck_D( IN := TRUE , PT := RobotLibraryParameter.INVALID_FRAMES_CHECK_TIMEOUT);

// Check Frame is valid : 
// ----------------------
// ST-FIX F66: an invalid frame is counted and not processed (spec 5.6.6.2)
_frameInvalid := ( _lifeSignHeader <> _lifeSignFooter );
IF ( _frameInvalid )
THEN
  AxesGroup.State.InvalidFrames := AxesGroup.State.InvalidFrames + 1;
END_IF


// Check timeout for invalid frame message
IF ( _invalidFrameCounterCheck_D.Q )
THEN
  // reset timer
 _invalidFrameCounterCheck_D( IN := FALSE);
  
  // compare invalid frame(s) counter
  IF ( AxesGroup.State.InvalidFrames <> _lastInvalidFrames)
  THEN
    // store last invalid frame(s) counter value
   _lastInvalidFrames := AxesGroup.State.InvalidFrames;
    // Create log entry
    CreateLogMessagePara1 ( Timestamp   := SystemTime,
                            MessageType := MessageType.CMD,
                            Severity    := Severity.WARNING,
                            MessageCode := 0,
                            MessageText := 'Detected invalid frames {1} in total',
                            Para1       :=  UDINT_TO_STRING(AxesGroup.State.InvalidFrames));
  END_IF
END_IF


// Reset invalid frames counter with rising edge of group reset
IF ( AxesGroup.State.GroupReset_R.Q)
THEN
  AxesGroup.State.InvalidFrames := 0;
             _lastInvalidFrames := 0;
 
  // Create log entry
  CreateLogMessage ( Timestamp   := SystemTime,
                     MessageType := MessageType.CMD,
                     Severity    := Severity.INFO,
                     MessageCode := 0,
                     MessageText := 'Reset invalid frames counter by executing GroupReset');
END_IF
                
                
END_METHOD

METHOD PRIVATE HandleLifeSign
VAR_IN_OUT
  /// Robot assignment of function
  AxesGroup    : AxesGroup;
END_VAR 
VAR_INST
  /// flag for 1st cycle
 _first : BOOL := TRUE;
END_VAR
                  IF ( _first ) OR ( NOT Enable ) 
THEN
  // init LifeSign 
  AxesGroup.Cyclic.PlcToRob.LifeSign := 0;
  // reset first flag
 _first := FALSE;
  // prevent inc LifeSign in the 1st cycle (Code below)
  RETURN;
END_IF


AxesGroup.Cyclic.PlcToRob.LifeSign := AxesGroup.Cyclic.PlcToRob.LifeSign + 1;
  
IF ( AxesGroup.Cyclic.PlcToRob.LifeSign > 15 )
THEN
  AxesGroup.Cyclic.PlcToRob.LifeSign := 1; // 0 is only in the very 1st cycle to indicate the system start in logging
END_IF


IF ( Enable ) AND ( _alive_F.Q ) 
THEN
  // Reset initialized flag
  Initialized := FALSE;
  // Reset Synchronized flag
  Synchronized := FALSE;
  
  // Set error 
  SetError( ErrorID := RobotLibraryErrorIdEnum.ERR_LIFESIGN_TIMEOUT_0x80A5 (* ST-FIX F65: lifesign timeout, table 7-2 *), Overwrite := TRUE );  
  // Create log entry
  CreateLogMessage ( Timestamp   := SystemTime,
                     MessageType := MessageType.CMD,
                     Severity    := Severity.FATAL_ERROR,
                     MessageCode := 0,
                     MessageText := 'LifeSign timeout -> Reinitialization required !');
END_IF

// Reset connection lost error
IF ( NOT Enable ) AND ( _aliveBit ) AND ( ErrorID = RobotLibraryErrorIdEnum.ERR_LIFESIGN_TIMEOUT_0x80A5 (* ST-FIX F65: lifesign timeout, table 7-2 *) )
THEN
  ErrorID := 0;
END_IF
                
                
END_METHOD

METHOD HandleLogMessagesAck
VAR_IN_OUT
   /// Robot assignment of function
  AxesGroup : AxesGroup;
END_VAR
                  IF ( _readMessages.Enabled )  
THEN
  // Set Message ID as Acknowlege ID  
 _readMessages.ParCmd.MsgID := _readMessages.OutCmd.MsgId;  
ELSE
  // Reset Acknowlege ID  
 _readMessages.ParCmd.MsgID := 0;
END_IF 



(*

IF (( _readMessages.Enabled           ) AND 
    ( _readMessages.OutCmd.MsgId > 0  ))  
THEN
  // Check if message has been entered into the message log ?   
  IF ( AxesGroup.MessageLog.CheckMessageCodePresent(_readMessages.OutCmd.ErrorCode ))
  THEN
    // Set Message ID as Acknowlege ID  
   _readMessages.ParCmd.MsgID := _readMessages.OutCmd.MsgId;  
	END_IF    
END_IF

*)
                
END_METHOD

METHOD PRIVATE HandleSeqAck
VAR_IN_OUT
   /// Robot assignment of function
  AxesGroup    : AxesGroup;
END_VAR 
VAR
  /// internal index for loops
 _idx : DINT;
END_VAR
                  // ST-FIX F63: Seq/Ack of one or two telegram sequences (spec 5.6.5.3, Fig. 5-206 ... 5-208):
//  - two sequences start with the Seq numbers 0 and 1
//  - the sequence with the lower Ack is handled first; its next Seq number is the number of the
//    other sequence + 1 (one common counter, the sequences alternate)
//  - ST-FIX F56: 254 -> 1, 0 only on the first exchange
IF ( _parCfg.Com.TwoSequences )
THEN
  AxesGroup.State.SequenceCountSend := 1;
ELSE
  AxesGroup.State.SequenceCountSend := 0;
END_IF

IF (NOT Enable)
THEN
  AxesGroup.State.CurrentSEQ[0] := 0;
  AxesGroup.State.CurrentSEQ[1] := DINT_TO_UINT(AxesGroup.State.SequenceCountSend);
END_IF

FOR _idx := 0 TO AxesGroup.State.SequenceCountSend
DO
  AxesGroup.State.CurrentAck[_idx] := Telegram.RobToPlc.Sequence[_idx].Header.SEQ_ACK;
END_FOR

  // ST-FIX F63: the sequence with the lower number first (Fig. 5-207/5-208), numbers wrap 254 -> 1
  _seqSendFirst := 0;
  IF ( AxesGroup.State.SequenceCountSend = 1 )
  THEN
    _seqDiff := UINT_TO_DINT(AxesGroup.State.CurrentAck[0]) - UINT_TO_DINT(AxesGroup.State.CurrentAck[1]);
    IF ( _seqDiff < 0 )
    THEN
      _seqDiff := _seqDiff + 254;
    END_IF
    IF ( _seqDiff > 0 ) AND ( _seqDiff < 127 )
    THEN
      _seqSendFirst := 1;
    END_IF
  END_IF

FOR _seqOrderIdx := 0 TO AxesGroup.State.SequenceCountSend
DO
  IF ( _seqOrderIdx = 0 )
  THEN
    _idx := _seqSendFirst;
  ELSE
    _idx := 1 - _seqSendFirst;
  END_IF

  // Check Seq/Ack :
  // ----------------------
  IF ( AxesGroup.State.CurrentAck[_idx] = AxesGroup.State.CurrentSEQ[_idx] )
  THEN
    _seqNext := AxesGroup.State.CurrentSEQ[AxesGroup.State.SequenceCountSend - _idx] + 1;
    IF ( _seqNext >= 255 )
    THEN
      _seqNext := 1;
    END_IF
    AxesGroup.State.CurrentSEQ[_idx] := _seqNext;
    AxesGroup.State.NewSEQ[_idx]     := TRUE;
  END_IF
END_FOR

// order in which the sequences are filled: lower Seq number first
// ST-FIX F63: the sequence with the lower number first (Fig. 5-207/5-208), numbers wrap 254 -> 1
_seqSendFirst := 0;
IF ( AxesGroup.State.SequenceCountSend = 1 )
THEN
  _seqDiff := UINT_TO_DINT(AxesGroup.State.CurrentSEQ[0]) - UINT_TO_DINT(AxesGroup.State.CurrentSEQ[1]);
  IF ( _seqDiff < 0 )
  THEN
    _seqDiff := _seqDiff + 254;
  END_IF
  IF ( _seqDiff > 0 ) AND ( _seqDiff < 127 )
  THEN
    _seqSendFirst := 1;
  END_IF
END_IF

// ST-FIX F65: telegram sequence timeout (spec 5.6.5.3/5.6.6.2: no new Seq number for
// 4 x LifeSignTimeOut while initialized) -> 16#80A8, reinitialization required
_seqAckTimeout( IN := Initialized AND NOT ( AxesGroup.State.NewSEQ[0] OR AxesGroup.State.NewSEQ[1] ),
                PT := 4 * ParCfg.Com.LifeSignTimeOut + ParCfg.Plc.CycleTime );
IF ( _seqAckTimeout.Q )
THEN
  Initialized  := FALSE;
  Synchronized := FALSE;
  SetError( ErrorID := RobotLibraryErrorIdEnum.ERR_TELEGRAM_SEQ_TIMEOUT_0x80A8 (* ST-FIX F180: correct name *), Overwrite := TRUE );
  CreateLogMessage ( Timestamp   := SystemTime,
                     MessageType := MessageType.CMD,
                     Severity    := Severity.FATAL_ERROR,
                     MessageCode := 0,
                     MessageText := 'Telegram sequence timeout -> Reinitialization required !');
END_IF
                
END_METHOD

METHOD PROTECTED HandleSync
VAR_IN_OUT
   /// Robot assignment of function
  AxesGroup : AxesGroup;
  /// ToolData stored on PLC.For more information refer to 5.5.6.4
  ToolData          : ARRAY[*] OF Tool;
  /// LoadData stored on PLC.For more information refer to 5.5.6.4
  FrameData         : ARRAY[*] OF Frame;
  /// LoadData stored on PLC.For more information refer to 5.5.6.4
  LoadData          : ARRAY[*] OF Load;
  /// Work areas stored on PLC. For more information refer to 5.5.8
  WorkAreas         : ARRAY[*] OF RobotWorkArea;
  /// Software limits stored on PLC
  SWLimits          : SWLimits;
  /// Default dynamics stored on PLC. For more information refer to 5.5.7
  DefaultDynamics   : DefaultDynamics;
  /// Reference dynamics stored on PLC. For more information refer to 5.5.7
  ReferenceDynamics : ReferenceDynamics;
END_VAR 

VAR
  /// flag that indicates at least any iten has enabled synchronisation
 _dataEnableSyncAny        : BOOL; 
  /// flag that indicates that the frame datas are synchronized or deactivated 
 _inSyncFrameOk            : BOOL;      
  /// flag that indicates that the tool datas are synchronized or deactivated 
 _inSyncToolOk             : BOOL;     
  /// flag that indicates that the load datas are synchronized or deactivated 
 _inSyncLoadOk             : BOOL;     
  /// flag that indicates that the work areas are synchronized or deactivated 
 _inSyncWorkAreaOk         : BOOL;
  /// flag that indicates that the SW limits are synchronized or deactivated 
 _inSyncSwLimitsOk         : BOOL;
  /// flag that indicates that the default dynamice are synchronized or deactivated 
 _inSyncDefaultDynamicOk   : BOOL;
  /// flag that indicates that the reference dynamice are synchronized or deactivated 
 _InSyncReferenceDynamicOk : BOOL;
END_VAR
                  HandleSyncToolData              ( AxesGroup := AxesGroup, ToolData          := ToolData);
HandleSyncFrameData             ( AxesGroup := AxesGroup, FrameData         := FrameData);
HandleSyncLoadData              ( AxesGroup := AxesGroup, LoadData          := LoadData);
HandleSyncRobotDefaultDynamics  ( AxesGroup := AxesGroup, DefaultDynamics   := DefaultDynamics);
HandleSyncRobotReferenceDynamics( AxesGroup := AxesGroup, ReferenceDynamics := ReferenceDynamics);
HandleSyncRobotSWLimits         ( AxesGroup := AxesGroup, SwLimits          := SwLimits);
// ST-FIX F13: HandleSyncToolData was called a second time here
HandleSyncWorkArea              ( AxesGroup := AxesGroup, WorkAreas         := WorkAreas);


// check any synchronisation activated ?
_dataEnableSyncAny :=        ((     AxesGroup.State.DataEnableSync.EnableSyncFrame             )  OR
                              (     AxesGroup.State.DataEnableSync.EnableSyncTool              )  OR
                              (     AxesGroup.State.DataEnableSync.EnableSyncLoad              )  OR
                              (     AxesGroup.State.DataEnableSync.EnableSyncWorkArea          )  OR
                              (     AxesGroup.State.DataEnableSync.EnableSyncSWLimits          )  OR
                              (     AxesGroup.State.DataEnableSync.EnableSyncDefaultDynamics   )  OR
                              (     AxesGroup.State.DataEnableSync.EnableSyncReferenceDynamics ));
                       
_inSyncFrameOk :=            ((     AxesGroup.State.SyncStatePlc     .InSync.Frame             )  AND 
                              (     AxesGroup.State.SyncStateRc      .InSync.Frame             )) OR
                              ( NOT AxesGroup.State.DataEnableSync.EnableSyncFrame ) OR // ST-FIX F24: not supported by the RC
( AxesGroup.State.Initialized AND NOT ( AxesGroup.State.RobotData.RCSupportedFunctions.ReadFrameData AND AxesGroup.State.RobotData.RCSupportedFunctions.WriteFrameData ));
                                                                                       
_inSyncToolOk :=             ((     AxesGroup.State.SyncStatePlc     .InSync.Tool              )  AND 
                              (     AxesGroup.State.SyncStateRc      .InSync.Tool              )) OR
                              ( NOT AxesGroup.State.DataEnableSync.EnableSyncTool ) OR // ST-FIX F24: not supported by the RC
( AxesGroup.State.Initialized AND NOT ( AxesGroup.State.RobotData.RCSupportedFunctions.ReadToolData AND AxesGroup.State.RobotData.RCSupportedFunctions.WriteToolData )); 
                                                                                           
_inSyncLoadOk :=             ((     AxesGroup.State.SyncStatePlc     .InSync.Load              )  AND 
                              (     AxesGroup.State.SyncStateRc      .InSync.Load              )) OR
                              ( NOT AxesGroup.State.DataEnableSync.EnableSyncLoad ) OR // ST-FIX F24: not supported by the RC
( AxesGroup.State.Initialized AND NOT ( AxesGroup.State.RobotData.RCSupportedFunctions.ReadLoadData AND AxesGroup.State.RobotData.RCSupportedFunctions.WriteLoadData )); 
                                                                                           
_inSyncWorkAreaOk :=         ((     AxesGroup.State.SyncStatePlc     .InSync.WorkArea          )  AND 
                              (     AxesGroup.State.SyncStateRc      .InSync.WorkArea          )) OR
                              ( NOT AxesGroup.State.DataEnableSync.EnableSyncWorkArea ) OR // ST-FIX F24: not supported by the RC
( AxesGroup.State.Initialized AND NOT ( AxesGroup.State.RobotData.RCSupportedFunctions.ReadWorkArea AND AxesGroup.State.RobotData.RCSupportedFunctions.WriteWorkArea )); 
                                                                                           
_inSyncSwLimitsOk :=         ((     AxesGroup.State.SyncStatePlc    .InSync.SwLimits           )  AND 
                              (     AxesGroup.State.SyncStateRc      .InSync.SwLimits          )) OR
                              ( NOT AxesGroup.State.DataEnableSync.EnableSyncSwLimits ) OR // ST-FIX F24: not supported by the RC
( AxesGroup.State.Initialized AND NOT ( AxesGroup.State.RobotData.RCSupportedFunctions.ReadRobotSWLimits AND AxesGroup.State.RobotData.RCSupportedFunctions.WriteRobotSWLimits )); 
                       
_inSyncDefaultDynamicOk :=   ((     AxesGroup.State.SyncStatePlc     .InSync.DefaultDynamics   )  AND 
                              (     AxesGroup.State.SyncStateRc      .InSync.DefaultDynamics   )) OR
                              ( NOT AxesGroup.State.DataEnableSync.EnableSyncDefaultDynamics ) OR // ST-FIX F24: not supported by the RC
( AxesGroup.State.Initialized AND NOT ( AxesGroup.State.RobotData.RCSupportedFunctions.ReadRobotDefaultDynamics AND AxesGroup.State.RobotData.RCSupportedFunctions.WriteRobotDefaultDynamics )); 

_inSyncReferenceDynamicOk := ((     AxesGroup.State.SyncStatePlc     .InSync.ReferenceDynamics )  AND 
                              (     AxesGroup.State.SyncStateRc      .InSync.ReferenceDynamics )) OR
                              ( NOT AxesGroup.State.DataEnableSync.EnableSyncReferenceDynamics ) OR // ST-FIX F24: not supported by the RC
( AxesGroup.State.Initialized AND NOT ( AxesGroup.State.RobotData.RCSupportedFunctions.ReadRobotReferenceDynamics AND AxesGroup.State.RobotData.RCSupportedFunctions.WriteRobotReferenceDynamics )); 
                       
                       
Synchronized := (( _inSyncFrameOk            ) AND      
                 ( _inSyncToolOk             ) AND    
                 ( _inSyncLoadOk             ) AND     
                 ( _inSyncWorkAreaOk         ) AND     
                 ( _inSyncSwLimitsOk         ) AND     
                 ( _inSyncDefaultDynamicOk   ) AND     
                 ( _InSyncReferenceDynamicOk ) AND            
                 ( _dataEnableSyncAny        ));                                                                                                                                                      


// Update exchange configuration parameter
_exchangeConfiguration.ParCmd.DataInSync.FramesInSync            := AxesGroup.State.SyncStatePlc.InSync.Frame;                // OR ( NOT AxesGroup.State.DataEnableSync.EnableSyncFrame            );
_exchangeConfiguration.ParCmd.DataInSync.ToolsInSync             := AxesGroup.State.SyncStatePlc.InSync.Tool;                 // OR ( NOT AxesGroup.State.DataEnableSync.EnableSyncTool             );
_exchangeConfiguration.ParCmd.DataInSync.LoadsInSync             := AxesGroup.State.SyncStatePlc.InSync.Load;                 // OR ( NOT AxesGroup.State.DataEnableSync.EnableSyncLoad             );
_exchangeConfiguration.ParCmd.DataInSync.WorkAreasInSync         := AxesGroup.State.SyncStatePlc.InSync.WorkArea;             // OR ( NOT AxesGroup.State.DataEnableSync.EnableSyncWorkArea         );
_exchangeConfiguration.ParCmd.DataInSync.SoftwareLimitsInSync    := AxesGroup.State.SyncStatePlc.InSync.SwLimits;             // OR ( NOT AxesGroup.State.DataEnableSync.EnableSyncSWLimits         );
_exchangeConfiguration.ParCmd.DataInSync.DefaultDynamicsInSync   := AxesGroup.State.SyncStatePlc.InSync.DefaultDynamics;      // OR ( NOT AxesGroup.State.DataEnableSync.EnableSyncDefaultDynamics  );
_exchangeConfiguration.ParCmd.DataInSync.ReferenceDynamicsInSync := AxesGroup.State.SyncStatePlc.InSync.ReferenceDynamics;    // OR ( NOT AxesGroup.State.DataEnableSync.EnableSyncReferenceDynamics);
                
                
END_METHOD

